               //BUFFER CONVEYOR LEVEL 5 - CONVEYOR 2
               "Control_DB".LCnv_Sys[3].Cnv_Level[5].Cnv2.Inputs.Left := NOT "C3205 - SENSOR CNV LEFT (FWD)";
               "Control_DB".LCnv_Sys[3].Cnv_Level[5].Cnv2.Inputs.Lpd1 := NOT "C3205 - SENSOR CNV LEFT (PALLET DETECT 1)";
               "Control_DB".LCnv_Sys[3].Cnv_Level[5].Cnv2.Inputs.Lpd2 := NOT "C3205 - SENSOR CNV LEFT (PALLET DETECT 2)";
               "Control_DB".LCnv_Sys[3].Cnv_Level[5].Cnv2.Inputs.Right := NOT "C3205 - SENSOR CNV RIGHT (BWD)";
               "Control_DB".LCnv_Sys[3].Cnv_Level[5].Cnv2.Inputs.Rpd1 := NOT "C3205 - SENSOR CNV RIGHT (PALLET DETECT 1)";
               "Control_DB".LCnv_Sys[3].Cnv_Level[5].Cnv2.Inputs.Rpd2 := NOT "C3205 - SENSOR CNV RIGHT (PALLET DETECT 2)";
               "Control_DB".LCnv_Sys[3].Cnv_Level[5].Cnv2.Inputs.Sdetect1 := NOT "C3205 - SHUTTLE IN POSITION 1";
               "Control_DB".LCnv_Sys[3].Cnv_Level[5].Cnv2.Inputs.Sdetect2 := NOT "C3205 - SHUTTLE IN POSITION 2";
               "Control_DB".LCnv_Sys[3].Cnv_Level[5].Cnv2.Safety_Stop_Cnrl.Inputs.DP_Extended := "C3205 - SENSOR SAFETY PIN1 UP";
               "Control_DB".LCnv_Sys[3].Cnv_Level[5].Cnv2.Safety_Stop_Cnrl.Inputs.DP_Retracted := "C3205 - SENSOR SAFETY PIN1 DOWN";

               "Control_DB".LCnv_Sys[3].Cnv_Level[5].Cnv2.Inputs.VFD_Status := "C3205_StatusWord";
               "Control_DB".LCnv_Sys[3].Cnv_Level[5].Cnv2.Inputs.VFD_ActualCurrent := WORD_TO_INT("C3205_ActualCurrent");
               "Control_DB".LCnv_Sys[3].Cnv_Level[5].Cnv2.Inputs.VFD_Speed_Actual := WORD_TO_INT("C3205_ActualSpeed");
               "Control_DB".LCnv_Sys[3].Cnv_Level[5].Cnv2.Inputs.VFD_ActualTorque := WORD_TO_INT("C3205_ActualTorque");
           END_REGION

           REGION LEVEL 6
               //BUFFER CONVEYOR LEVEL 6 - CONVEYOR 1
               "Control_DB".LCnv_Sys[3].Cnv_Level[6].Cnv1.Inputs.Left := NOT "C3106 - SENSOR CNV LEFT (FWD)";
               "Control_DB".LCnv_Sys[3].Cnv_Level[6].Cnv1.Inputs.Lpd1 := NOT "C3106 - SENSOR CNV LEFT (PALLET DETECT 1)";
               "Control_DB".LCnv_Sys[3].Cnv_Level[6].Cnv1.Inputs.Lpd2 := NOT "C3106 - SENSOR CNV LEFT (PALLET DETECT 2)";
               "Control_DB".LCnv_Sys[3].Cnv_Level[6].Cnv1.Inputs.Right := NOT "C3106 - SENSOR CNV RIGHT (BWD)";
               "Control_DB".LCnv_Sys[3].Cnv_Level[6].Cnv1.Inputs.Rpd1 := NOT "C3106 - SENSOR CNV RIGHT (PALLET DETECT 1)";
               "Control_DB".LCnv_Sys[3].Cnv_Level[6].Cnv1.Inputs.Rpd2 := NOT "C3106 - SENSOR CNV RIGHT (PALLET DETECT 2)";
               "Control_DB".LCnv_Sys[3].Cnv_Level[6].Cnv1.Inputs.Sdetect1 := NOT "C3106 - SHUTTLE IN POSITION 1";
               "Control_DB".LCnv_Sys[3].Cnv_Level[6].Cnv1.Inputs.Sdetect2 := NOT "C3106 - SHUTTLE IN POSITION 2";
               "Control_DB".LCnv_Sys[3].Cnv_Level[6].Cnv1.Safety_Stop_Cnrl.Inputs.DP_Extended := "C3106 - SENSOR SAFETY PIN1 UP";
               "Control_DB".LCnv_Sys[3].Cnv_Level[6].Cnv1.Safety_Stop_Cnrl.Inputs.DP_Retracted := "C3106 - SENSOR SAFETY PIN1 DOWN";

               "Control_DB".LCnv_Sys[3].Cnv_Level[6].Cnv1.Inputs.VFD_Status := "C3106_StatusWord";
               "Control_DB".LCnv_Sys[3].Cnv_Level[6].Cnv1.Inputs.VFD_ActualCurrent := WORD_TO_INT("C3106_ActualCurrent");
               "Control_DB".LCnv_Sys[3].Cnv_Level[6].Cnv1.Inputs.VFD_Speed_Actual := WORD_TO_INT("C3106_ActualSpeed");
               "Control_DB".LCnv_Sys[3].Cnv_Level[6].Cnv1.Inputs.VFD_ActualTorque := WORD_TO_INT("C3106_ActualTorque");

               //BUFFER CONVEYOR LEVEL 6 - CONVEYOR 2
               "Control_DB".LCnv_Sys[3].Cnv_Level[6].Cnv2.Inputs.Left := NOT "C3206 - SENSOR CNV LEFT (FWD)";
               "Control_DB".LCnv_Sys[3].Cnv_Level[6].Cnv2.Inputs.Lpd1 := NOT "C3206 - SENSOR CNV LEFT (PALLET DETECT 1)";
               "Control_DB".LCnv_Sys[3].Cnv_Level[6].Cnv2.Inputs.Lpd2 := NOT "C3206 - SENSOR CNV LEFT (PALLET DETECT 2)";
               "Control_DB".LCnv_Sys[3].Cnv_Level[6].Cnv2.Inputs.Right := NOT "C3206 - SENSOR CNV RIGHT (BWD)";
               "Control_DB".LCnv_Sys[3].Cnv_Level[6].Cnv2.Inputs.Rpd1 := NOT "C3206 - SENSOR CNV RIGHT (PALLET DETECT 1)";
               "Control_DB".LCnv_Sys[3].Cnv_Level[6].Cnv2.Inputs.Rpd2 := NOT "C3206 - SENSOR CNV RIGHT (PALLET DETECT 2)";
               "Control_DB".LCnv_Sys[3].Cnv_Level[6].Cnv2.Inputs.Sdetect1 := NOT "C3206 - SHUTTLE IN POSITION 1";
               "Control_DB".LCnv_Sys[3].Cnv_Level[6].Cnv2.Inputs.Sdetect2 := NOT "C3206 - SHUTTLE IN POSITION 2";
               "Control_DB".LCnv_Sys[3].Cnv_Level[6].Cnv2.Safety_Stop_Cnrl.Inputs.DP_Extended := "C3206 - SENSOR SAFETY PIN1 UP";
               "Control_DB".LCnv_Sys[3].Cnv_Level[6].Cnv2.Safety_Stop_Cnrl.Inputs.DP_Retracted := "C3206 - SENSOR SAFETY PIN1 DOWN";

               "Control_DB".LCnv_Sys[3].Cnv_Level[6].Cnv2.Inputs.VFD_Status := "C3206_StatusWord";
               "Control_DB".LCnv_Sys[3].Cnv_Level[6].Cnv2.Inputs.VFD_ActualCurrent := WORD_TO_INT("C3206_ActualCurrent");
               "Control_DB".LCnv_Sys[3].Cnv_Level[6].Cnv2.Inputs.VFD_Speed_Actual := WORD_TO_INT("C3206_ActualSpeed");
               "Control_DB".LCnv_Sys[3].Cnv_Level[6].Cnv2.Inputs.VFD_ActualTorque := WORD_TO_INT("C3206_ActualTorque");
           END_REGION

           REGION LEVEL 7
               //BUFFER CONVEYOR LEVEL 7 - CONVEYOR 1
               "Control_DB".LCnv_Sys[3].Cnv_Level[7].Cnv1.Inputs.Left := NOT "C3107 - SENSOR CNV LEFT (FWD)";
               "Control_DB".LCnv_Sys[3].Cnv_Level[7].Cnv1.Inputs.Lpd1 := NOT "C3107 - SENSOR CNV LEFT (PALLET DETECT 1)";
               "Control_DB".LCnv_Sys[3].Cnv_Level[7].Cnv1.Inputs.Lpd2 := NOT "C3107 - SENSOR CNV LEFT (PALLET DETECT 2)";
               "Control_DB".LCnv_Sys[3].Cnv_Level[7].Cnv1.Inputs.Right := NOT "C3107 - SENSOR CNV RIGHT (BWD)";
               "Control_DB".LCnv_Sys[3].Cnv_Level[7].Cnv1.Inputs.Rpd1 := NOT "C3107 - SENSOR CNV RIGHT (PALLET DETECT 1)";
               "Control_DB".LCnv_Sys[3].Cnv_Level[7].Cnv1.Inputs.Rpd2 := NOT "C3107 - SENSOR CNV RIGHT (PALLET DETECT 2)";
               "Control_DB".LCnv_Sys[3].Cnv_Level[7].Cnv1.Inputs.Sdetect1 := NOT "C3107 - SHUTTLE IN POSITION 1";
               "Control_DB".LCnv_Sys[3].Cnv_Level[7].Cnv1.Inputs.Sdetect2 := NOT "C3107 - SHUTTLE IN POSITION 2";
               "Control_DB".LCnv_Sys[3].Cnv_Level[7].Cnv1.Safety_Stop_Cnrl.Inputs.DP_Extended := "C3107 - SENSOR SAFETY PIN1 UP";
               "Control_DB".LCnv_Sys[3].Cnv_Level[7].Cnv1.Safety_Stop_Cnrl.Inputs.DP_Retracted := "C3107 - SENSOR SAFETY PIN1 DOWN";

               "Control_DB".LCnv_Sys[3].Cnv_Level[7].Cnv1.Inputs.VFD_Status := "C3107_StatusWord";
               "Control_DB".LCnv_Sys[3].Cnv_Level[7].Cnv1.Inputs.VFD_ActualCurrent := WORD_TO_INT("C3107_ActualCurrent");
               "Control_DB".LCnv_Sys[3].Cnv_Level[7].Cnv1.Inputs.VFD_Speed_Actual := WORD_TO_INT("C3107_ActualSpeed");
               "Control_DB".LCnv_Sys[3].Cnv_Level[7].Cnv1.Inputs.VFD_ActualTorque := WORD_TO_INT("C3107_ActualTorque");

               //BUFFER CONVEYOR LEVEL 7 - CONVEYOR 2
               "Control_DB".LCnv_Sys[3].Cnv_Level[7].Cnv2.Inputs.Left := NOT "C3207 - SENSOR CNV LEFT (FWD)";
               "Control_DB".LCnv_Sys[3].Cnv_Level[7].Cnv2.Inputs.Lpd1 := NOT "C3207 - SENSOR CNV LEFT (PALLET DETECT 1)";
               "Control_DB".LCnv_Sys[3].Cnv_Level[7].Cnv2.Inputs.Lpd2 := NOT "C3207 - SENSOR CNV LEFT (PALLET DETECT 2)";
               "Control_DB".LCnv_Sys[3].Cnv_Level[7].Cnv2.Inputs.Right := NOT "C3207 - SENSOR CNV RIGHT (BWD)";
               "Control_DB".LCnv_Sys[3].Cnv_Level[7].Cnv2.Inputs.Rpd1 := NOT "C3207 - SENSOR CNV RIGHT (PALLET DETECT 1)";
               "Control_DB".LCnv_Sys[3].Cnv_Level[7].Cnv2.Inputs.Rpd2 := NOT "C3207 - SENSOR CNV RIGHT (PALLET DETECT 2)";
               "Control_DB".LCnv_Sys[3].Cnv_Level[7].Cnv2.Inputs.Sdetect1 := NOT "C3207 - SHUTTLE IN POSITION 1";
               "Control_DB".LCnv_Sys[3].Cnv_Level[7].Cnv2.Inputs.Sdetect2 := NOT "C3207 - SHUTTLE IN POSITION 2";
               "Control_DB".LCnv_Sys[3].Cnv_Level[7].Cnv2.Safety_Stop_Cnrl.Inputs.DP_Extended := "C3207 - SENSOR SAFETY PIN1 UP";
               "Control_DB".LCnv_Sys[3].Cnv_Level[7].Cnv2.Safety_Stop_Cnrl.Inputs.DP_Retracted := "C3207 - SENSOR SAFETY PIN1 DOWN";

               "Control_DB".LCnv_Sys[3].Cnv_Level[7].Cnv2.Inputs.VFD_Status := "C3207_StatusWord";
               "Control_DB".LCnv_Sys[3].Cnv_Level[7].Cnv2.Inputs.VFD_ActualCurrent := WORD_TO_INT("C3207_ActualCurrent");
               "Control_DB".LCnv_Sys[3].Cnv_Level[7].Cnv2.Inputs.VFD_Speed_Actual := WORD_TO_INT("C3207_ActualSpeed");
               "Control_DB".LCnv_Sys[3].Cnv_Level[7].Cnv2.Inputs.VFD_ActualTorque := WORD_TO_INT("C3207_ActualTorque");
           END_REGION

           REGION LEVEL 8
               //BUFFER CONVEYOR LEVEL 8 - CONVEYOR 1
               "Control_DB".LCnv_Sys[3].Cnv_Level[8].Cnv1.Inputs.Left := NOT "C3108 - SENSOR CNV LEFT (FWD)";
               "Control_DB".LCnv_Sys[3].Cnv_Level[8].Cnv1.Inputs.Lpd1 := NOT "C3108 - SENSOR CNV LEFT (PALLET DETECT 1)";
               "Control_DB".LCnv_Sys[3].Cnv_Level[8].Cnv1.Inputs.Lpd2 := NOT "C3108 - SENSOR CNV LEFT (PALLET DETECT 2)";
               "Control_DB".LCnv_Sys[3].Cnv_Level[8].Cnv1.Inputs.Right := NOT "C3108 - SENSOR CNV RIGHT (BWD)";
               "Control_DB".LCnv_Sys[3].Cnv_Level[8].Cnv1.Inputs.Rpd1 := NOT "C3108 - SENSOR CNV RIGHT (PALLET DETECT 1)";
               "Control_DB".LCnv_Sys[3].Cnv_Level[8].Cnv1.Inputs.Rpd2 := NOT "C3108 - SENSOR CNV RIGHT (PALLET DETECT 2)";
               "Control_DB".LCnv_Sys[3].Cnv_Level[8].Cnv1.Inputs.Sdetect1 := NOT "C3108 - SHUTTLE IN POSITION 1";
               "Control_DB".LCnv_Sys[3].Cnv_Level[8].Cnv1.Inputs.Sdetect2 := NOT "C3108 - SHUTTLE IN POSITION 2";
               "Control_DB".LCnv_Sys[3].Cnv_Level[8].Cnv1.Safety_Stop_Cnrl.Inputs.DP_Extended := "C3108 - SENSOR SAFETY PIN1 UP";
               "Control_DB".LCnv_Sys[3].Cnv_Level[8].Cnv1.Safety_Stop_Cnrl.Inputs.DP_Retracted := "C3108 - SENSOR SAFETY PIN1 DOWN";

               "Control_DB".LCnv_Sys[3].Cnv_Level[8].Cnv1.Inputs.VFD_Status := "C3108_StatusWord";
               "Control_DB".LCnv_Sys[3].Cnv_Level[8].Cnv1.Inputs.VFD_ActualCurrent := WORD_TO_INT("C3108_ActualCurrent");
               "Control_DB".LCnv_Sys[3].Cnv_Level[8].Cnv1.Inputs.VFD_Speed_Actual := WORD_TO_INT("C3108_ActualSpeed");
               "Control_DB".LCnv_Sys[3].Cnv_Level[8].Cnv1.Inputs.VFD_ActualTorque := WORD_TO_INT("C3108_ActualTorque");

               //BUFFER CONVEYOR LEVEL 8 - CONVEYOR 2
               "Control_DB".LCnv_Sys[3].Cnv_Level[8].Cnv2.Inputs.Left := NOT "C3208 - SENSOR CNV LEFT (FWD)";
               "Control_DB".LCnv_Sys[3].Cnv_Level[8].Cnv2.Inputs.Lpd1 := NOT "C3208 - SENSOR CNV LEFT (PALLET DETECT 1)";
               "Control_DB".LCnv_Sys[3].Cnv_Level[8].Cnv2.Inputs.Lpd2 := NOT "C3208 - SENSOR CNV LEFT (PALLET DETECT 2)";
               "Control_DB".LCnv_Sys[3].Cnv_Level[8].Cnv2.Inputs.Right := NOT "C3208 - SENSOR CNV RIGHT (BWD)";
               "Control_DB".LCnv_Sys[3].Cnv_Level[8].Cnv2.Inputs.Rpd1 := NOT "C3208 - SENSOR CNV RIGHT (PALLET DETECT 1)";
               "Control_DB".LCnv_Sys[3].Cnv_Level[8].Cnv2.Inputs.Rpd2 := NOT "C3208 - SENSOR CNV RIGHT (PALLET DETECT 2)";
               "Control_DB".LCnv_Sys[3].Cnv_Level[8].Cnv2.Inputs.Sdetect1 := NOT "C3208 - SHUTTLE IN POSITION 1";
               "Control_DB".LCnv_Sys[3].Cnv_Level[8].Cnv2.Inputs.Sdetect2 := NOT "C3208 - SHUTTLE IN POSITION 2";
               "Control_DB".LCnv_Sys[3].Cnv_Level[8].Cnv2.Safety_Stop_Cnrl.Inputs.DP_Extended := "C3208 - SENSOR SAFETY PIN1 UP";
               "Control_DB".LCnv_Sys[3].Cnv_Level[8].Cnv2.Safety_Stop_Cnrl.Inputs.DP_Retracted := "C3208 - SENSOR SAFETY PIN1 DOWN";

               "Control_DB".LCnv_Sys[3].Cnv_Level[8].Cnv2.Inputs.VFD_Status := "C3208_StatusWord";
               "Control_DB".LCnv_Sys[3].Cnv_Level[8].Cnv2.Inputs.VFD_ActualCurrent := WORD_TO_INT("C3208_ActualCurrent");
               "Control_DB".LCnv_Sys[3].Cnv_Level[8].Cnv2.Inputs.VFD_Speed_Actual := WORD_TO_INT("C3208_ActualSpeed");
               "Control_DB".LCnv_Sys[3].Cnv_Level[8].Cnv2.Inputs.VFD_ActualTorque := WORD_TO_INT("C3208_ActualTorque");
           END_REGION
       END_REGION

       REGION VTD
           "Control_DB".VTD_Sys[3].Inputs.Upper_Overtravel := "OVERTRAVEL UPPER LIMIT - CH1(3)";
           "Control_DB".VTD_Sys[3].Inputs.Upper_limit := "VTD3 UPPER LIMIT";
           "Control_DB".VTD_Sys[3].Inputs.Ultimate_SlowDown := "VTD3 ULTIMATE SLOWDOWN";
           "Control_DB".VTD_Sys[3].Inputs.Ultimate_Creep := "VTD3 ULTIMATE CREEP";
           "Control_DB".VTD_Sys[3].Inputs.Lower_Limit := "VTD3 LOWER LIMIT";
           "Control_DB".VTD_Sys[3].Inputs.Lower_Overtravel := "OVERTRAVEL LOWER LIMIT - CH1(3)";
           "Control_DB".VTD_Sys[3].Inputs.Level_Detect1 := "VTD3 LEVEL DETECT 1";
           "Control_DB".VTD_Sys[3].Inputs.Level_Detect2 := "VTD3 LEVEL DETECT 2";
           "Control_DB".VTD_Sys[3].Inputs.DP1_Extended := "VTD3 DOCKING PINS EXTENDED 1";
           "Control_DB".VTD_Sys[3].Inputs.DP2_Extended := "VTD3 DOCKING PINS EXTENDED 2";
           "Control_DB".VTD_Sys[3].Inputs.DP1_Retracted := "VTD3 DOCKING PINS RETRACTED 1";
           "Control_DB".VTD_Sys[3].Inputs.DP2_Retracted := "VTD3 DOCKING PINS RETRACTED 2";
           "Control_DB".VTD_Sys[3].Inputs.Chain_Slack_1 := NOT "Remote_Panel_DB_3".Chain_Slack_1_Filtered;
           "Control_DB".VTD_Sys[3].Inputs.Chain_Slack_2 := NOT "Remote_Panel_DB_3".Chain_Slack_2_Filtered;
           "Control_DB".VTD_Sys[3].Inputs.Chain_Slack_3 := NOT "Remote_Panel_DB_3".Chain_Slack_3_Filtered;
           "Control_DB".VTD_Sys[3].Inputs.Chain_Slack_4 := NOT "Remote_Panel_DB_3".Chain_Slack_4_Filtered;
           "Control_DB".VTD_Sys[3].Inputs.PushToEnter := "VTD3 PUSH TO ENTER VTD ZONE";
           "Control_DB".VTD_Sys[3].Inputs.PushToExit := "VTD3 PUSH TO EXIT VTD ZONE";

           "Control_DB".VTD_Sys[3].Inputs.VFD_Status := "VTD3_StatusWord";
           "Control_DB".VTD_Sys[3].Inputs.VFD_ActualCurrent := REAL_TO_INT(("VTD3_ActualCurrent" / 10) / 72.5);
           "Control_DB".VTD_Sys[3].Inputs.VFD_Speed_Actual := "VTD3_ActualSpeed";
           "Control_DB".VTD_Sys[3].Inputs.VFD_ActualTorque := WORD_TO_INT("VTD3_ActualTorque");

       END_REGION

       REGION ABSOLUTE ENCODER
           REGION DOCUMENTATION
               //STATUS---------------------------------------------------------------------------------------------------------------------
               //
               //Encoder state word 2 - INPUT WORD 1
               //
               // 15 … 12 Encoder’s Sign-OF-Life (NOT relevant)
               // 11, 10 Reserved
               // 9 Control requested 0 = No control BY the PLC requested 1 = Control BY the PLC requested
               // 8 … 0 Reserved

               //Sensor 1 state word - INPUT WORD 2
               //
               // 15 Encoder error Description 0 = No error 1 = Error The error code is output in G1_XIST2.
               // 14 Park mode activated 0 = Normal operation 1 = Park mode activated Feedback based on G1_STW bit 14: No output OF position data G1_XIST1 AND G1_XIST2
               // 13 Transmission OF absolute position value 0 = No transmission 1 = Position value is output in G1_XIST2
               // 12 Status OF the Preset function (set/shift OF home position executed) 0 = No Preset function active 1 = Preset function is run Feedback based on G1_STW bit 12:  
               // 11 Requirement OF error acknowledgement detected New position value is output in G1_XIST1 AND G1_XIST2. On conclusion OF the Preset function the bit is set TO 0. 0 = No RETURN acknowledgement OF Encoder error 1 = Requirement OF error acknowledgement detected Reaction TO bit 15 in the sensor control word 1 G1_STW is acknowledged (see Table 14)
               // 10 Reserved
               // 9 … 0 NOT supported

               //Position 1 - INPUT WORD 3 AND 4
               // "AE_Position_1_Scaled" := (*SCALE_X(MIN := "Settings_DB".VTD_Settings.VTD_Min_Height,
               //                                   VALUE := *)NORM_X(MIN := 0,
               //                                                   VALUE := (SHL(IN:="AE_Position_1", N:=2) * 0.00228881) (*- "AE_Offset"*),
               //                                                   MAX := 1073741824)(*,
               //                                   MAX := "Settings_DB".VTD_Settings.VTD_Max_Heigh)*);
               // "mm_per_pulse" := 401,5584 / 262144;
               // 
               //CONTROL---------------------------------------------------------------------------------------------------------------------
               //
               //Encoder control word 2 - OUTPUT WORD 1
               //
               // 15 … 12 Master’s Sign-OF-Life (NOT relevant)
               // 10 control BY PLC 0 = No control BY the PLC 1 = Control BY the PLC Enables the PLC BY using control words TO activate / deactivate encoder functions
               // 7 Fault acknowledge Error-buffer handling NOT supported
               // 11, 9, 8, 6 … 0 Reserved
               // "AE_Control_Word_1".%X10 := "AE_PLC_Control";
               // 
               //Sensor 1 control word - OUTPUT WORD 2-------------------------------------------------------------------------------------------
               //
               // 15 Acknowledging a sensor error Description 0 = Encoder error message NOT acknowledged BY PLC 1 = Encoder error message acknowledged BY the PLC
               // 14 Activate park mode 0 = Normal operation 1 = Activate park mode
               // 13 Request FOR the absolute position value 0 = No request 1 = Request BY the master Results in the cyclic output OF the position values in G1_XIST2
               // 12 Activate preset value (see note below) Defines that a configured preset value is used (see section 3.5 on page 24) 0 = Preset value is NOT activated 1 = Preset value is activated
               // 11 Preset mode Defines how a configured preset value is used 0 = Preset value is used as a new absolute value 1 = Preset value is added TO the previous value
               // 10 … 0 Reserved
               // "AE_Control_Word_2".%X15 := "VTD_Reset_HMI_Tags";
               // "AE_Control_Word_2".%X14 := "AE_Activate_ParkMode";
               // "AE_Control_Word_2".%X13 := "AE_Request_ABS_Value";
               // "AE_Control_Word_2".%X12 := "AE_Activate_Preset_Value";
               // "AE_Control_Word_2".%X11 := "AE_Preset_Mode";
           END_REGION

           //STATUS---------------------------------------------------------------------------------------------------------------------
           "Control_DB".VTD_Sys[3].Inputs.AE_Status_2 := "AE_Status_2(3)";
           //Position 1 - INPUT WORD 3 AND 4
           "Control_DB".VTD_Sys[3].Inputs.AE_Position_1 := REAL_TO_DINT(((((*1073741823 - reverse the direction*)
         (SHR(IN := "AE_Position_1(3)", N := 2))) - 31381317) * 0.0015318237304688 (*Mechanical relationship*)- 225511)(*Offset*));

           // Position 2 - INPUT WORD 5 AND 6
           "Control_DB".VTD_Sys[3].Inputs.AE_Position_2 := SHR(IN := "AE_Position_2(3)", N := 2);

           //Speed A - INPUT WORD 7
           "Control_DB".VTD_Sys[3].Inputs.AE_Speed := "AE_Speed(3)";
       END_REGION

       REGION LINEAR ENCODER
           "Control_DB".VTD_Sys[3].Inputs.LE_Position := "LE_X_Unsafe_Position(3)" / 10;
           "Control_DB".VTD_Sys[3].Inputs.LE_Speed := "LE_Speed(3)" * 100;
           "Control_DB".VTD_Sys[3].Inputs.LE_Status := "LE_Status(3)";
           "Control_DB".VTD_Sys[3].Inputs.LE_Warnings := "LE_Warnings(3)";
           REGION DOCUMENTATION
               //STATUS 
               //
               // 0 ERR - Error message (Error code in XP00– XP15); remaining bits = 0, see Error Codes
               // 1 NP - No position information/OUT (XP = 0, YP = 0, SP = 0)
               // 2 WRN - Warnings present, see Warning Module
               // 3 EV - Event present
               // 4 posdetected - Valid position information available

               //WARNINGS
               //
               // 0 WRN01 A code with non-PXV content was found.
               // 1 WRN02 the read head is too close TO the Data Matrix code tape.
               // 2 WRN03 the read head is too far from the Data Matrix code tape.
               // 3 WRN04 Y position too large. The sensor is just before OUT.
               // 4 WRN05 Y position is too small. The sensor is just before OUT.
               // 5 WRN06 the read head is rotated OR tilted in relation TO the Data Matrix code tape.
               // 6 WRN07 Low level OF code contrast.
               // 7 WRN08 Repair tape detected.
               // 8 WRN09 Temperature too high.
               // 9...15 Reserved

               //QUALITY GRADE
               //
               //The quality grades enable constant monitoring of the code tape and the camera along the entire
               //traverse distance. This enables you to detect and act upon potential damage or contamination
               //of the code tape and camera at the earliest stage possible during commissioning and normal
               //operation. As a result, this maximizes the overall functional reliability of your plant, and
               //it means you are able to immediately localize the issue in the case of a fault. Evaluations
               //are made using a scale of 1 to 6. The value 1 is the best possible read quality. A value greater
               //than 3 or worse requires the camera and its path to be inspected. The value 7 signifies "No position"
               //because no code was detected. An evaluation that indicates poor quality as the outcome can be due to
               //a misalignment or incorrect orientation, an incorrect measuring distance, or because the code tape has been affixed incorrectly
           END_REGION
       END_REGION

       REGION SICK BARCODE LECTORS
           IF "Control_DB".VTDBarcode_Station[3].Running AND "SICK_Lector_Control_DB_3".Result <> "Control_DB".VTDBarcode_Station[3].Barcode_Old THEN
               "Control_DB".VTD_Sys[3].Inputs."Barcode 1" := "SICK_Lector_Control_DB_3".Result;
               // "Control_DB".VTD_Control.Inputs."Barcode 2'" := SICK_Barcode_DB".Result;
               // "Control_DB".VTDBarcode_Station[3].Barcode_Old := "SICK_Lector_Control_DB_3".Result;
           ELSE
               "Control_DB".VTD_Sys[3].Inputs."Barcode 1" :=
               "Control_DB".VTD_Sys[3].Inputs."Barcode 2" := '';
           END_IF;

       END_REGION

       REGION VFD HARDWARE ID
           //Buffer conveyors 1
           "Settings_DB".LCnv_Sys[3].Cnv_Level[1].Cnv1.G120_Hardware_ID := "C3101~Drive_1~Standard_telegram_20__PZD-2_6";
           "Settings_DB".LCnv_Sys[3].Cnv_Level[2].Cnv1.G120_Hardware_ID := "C3102~Drive_1~Standard_telegram_20__PZD-2_6";
           "Settings_DB".LCnv_Sys[3].Cnv_Level[3].Cnv1.G120_Hardware_ID := "C3103~Drive_1~Standard_telegram_20__PZD-2_6";
           "Settings_DB".LCnv_Sys[3].Cnv_Level[4].Cnv1.G120_Hardware_ID := "C3104~Drive_1~Standard_telegram_20__PZD-2_6";
           "Settings_DB".LCnv_Sys[3].Cnv_Level[5].Cnv1.G120_Hardware_ID := "C3105~Drive_1~Standard_telegram_20__PZD-2_6";
           "Settings_DB".LCnv_Sys[3].Cnv_Level[6].Cnv1.G120_Hardware_ID := "C3106~Drive_1~Standard_telegram_20__PZD-2_6";
           "Settings_DB".LCnv_Sys[3].Cnv_Level[7].Cnv1.G120_Hardware_ID := "C3107~Drive_1~Standard_telegram_20__PZD-2_6";
           "Settings_DB".LCnv_Sys[3].Cnv_Level[8].Cnv1.G120_Hardware_ID := "C3108~Drive_1~Standard_telegram_20__PZD-2_6";

           //Buffer conveyors 2
           "Settings_DB".LCnv_Sys[3].Cnv_Level[1].Cnv2.G120_Hardware_ID := "C3201~Drive_1~Standard_telegram_20__PZD-2_6";
           "Settings_DB".LCnv_Sys[3].Cnv_Level[2].Cnv2.G120_Hardware_ID := "C3202~Drive_1~Standard_telegram_20__PZD-2_6";
           "Settings_DB".LCnv_Sys[3].Cnv_Level[3].Cnv2.G120_Hardware_ID := "C3203~Drive_1~Standard_telegram_20__PZD-2_6";
           "Settings_DB".LCnv_Sys[3].Cnv_Level[4].Cnv2.G120_Hardware_ID := "C3204~Drive_1~Standard_telegram_20__PZD-2_6";
           "Settings_DB".LCnv_Sys[3].Cnv_Level[5].Cnv2.G120_Hardware_ID := "C3205~Drive_1~Standard_telegram_20__PZD-2_6";
           "Settings_DB".LCnv_Sys[3].Cnv_Level[6].Cnv2.G120_Hardware_ID := "C3206~Drive_1~Standard_telegram_20__PZD-2_6";
           "Settings_DB".LCnv_Sys[3].Cnv_Level[7].Cnv2.G120_Hardware_ID := "C3207~Drive_1~Standard_telegram_20__PZD-2_6";
           "Settings_DB".LCnv_Sys[3].Cnv_Level[8].Cnv2.G120_Hardware_ID := "C3208~Drive_1~Standard_telegram_20__PZD-2_6";

           //Extractor conveyor
           "Settings_DB".ECnv_Sys[3].G120_Hardware_ID := "CVTD_3~Drive_1~Standard_telegram_20__PZD-2_6";

           //VTD
           "Settings_DB".VTD_Sys[3].G120_Hardware_ID := "VTD_3~DO_VECTOR_1~Standard_telegram_20__PZD-2_6";
       END_REGION
   END_REGION

   REGION SYSTEM 4
       REGION EXTRACTOR CONVEYOR
           "Control_DB".ECnv_Sys[4].Inputs.Left := "CVTD4 SENSOR CONVEYOR LEFT (FWD)";
           "Control_DB".ECnv_Sys[4].Inputs.Lpd1 := "CVTD4 SENSOR CONVEYOR LEFT (PALLET DETECT 1)";
           "Control_DB".ECnv_Sys[4].Inputs.Center := "CVTD4 SENSOR CONVEYOR CENTER";
           "Control_DB".ECnv_Sys[4].Inputs.Right := "CVTD4 SENSOR CONVEYOR RIGHT (BWD)";
           "Control_DB".ECnv_Sys[4].Inputs.Rpd1 := "CVTD4 SENSOR CONVEYOR RIGHT (PALLET DETECT 1)";

           "T_OH_Left_4".TOF(IN := "CVTD4 OVERHANG LEFT" OR NOT "Control_DB".VTD_Sys[4].Running,
                             PT := T#200ms);
           "Control_DB".ECnv_Sys[4].Inputs.Overhang_Left := "T_OH_Left_4".Q;

           "I_OH_Right_4".TOF(IN := "CVTD4 OVERHANG RIGHT" OR NOT "Control_DB".VTD_Sys[4].Running,
                              PT := T#200ms);
           "Control_DB".ECnv_Sys[4].Inputs.Overhang_Right := "I_OH_Right_4".Q;

           "Control_DB".ECnv_Sys[4].Inputs.VFD_Status := "CVTD4_StatusWord";
           "Control_DB".ECnv_Sys[4].Inputs.VFD_ActualCurrent := WORD_TO_INT("CVTD4_ActualCurrent");
           "Control_DB".ECnv_Sys[4].Inputs.VFD_Speed_Actual := WORD_TO_INT("CVTD4_ActualSpeed");
           "Control_DB".ECnv_Sys[4].Inputs.VFD_ActualTorque := WORD_TO_INT("CVTD4_ActualTorque");
       END_REGION

       REGION BUFFER CONVEYORS
           REGION LEVEL 1
               //BUFFER CONVEYOR LEVEL 1 - CONVEYOR 1
               "Control_DB".LCnv_Sys[4].Cnv_Level[1].Cnv1.Inputs.Left := NOT "C4101 - SENSOR CNV LEFT (FWD)";
               "Control_DB".LCnv_Sys[4].Cnv_Level[1].Cnv1.Inputs.Lpd1 := NOT "C4101 - SENSOR CNV LEFT (PALLET DETECT 1)";
               "Control_DB".LCnv_Sys[4].Cnv_Level[1].Cnv1.Inputs.Lpd2 := NOT "C4101 - SENSOR CNV LEFT (PALLET DETECT 2)";
               "Control_DB".LCnv_Sys[4].Cnv_Level[1].Cnv1.Inputs.Right := NOT "C4101 - SENSOR CNV RIGHT (BWD)";
               "Control_DB".LCnv_Sys[4].Cnv_Level[1].Cnv1.Inputs.Rpd1 := NOT "C4101 - SENSOR CNV RIGHT (PALLET DETECT 1)";
               "Control_DB".LCnv_Sys[4].Cnv_Level[1].Cnv1.Inputs.Rpd2 := NOT "C4101 - SENSOR CNV RIGHT (PALLET DETECT 2)";
               "Control_DB".LCnv_Sys[4].Cnv_Level[1].Cnv1.Inputs.Sdetect1 := NOT "C4101 - SHUTTLE IN POSITION 1";
               "Control_DB".LCnv_Sys[4].Cnv_Level[1].Cnv1.Inputs.Sdetect2 := NOT "C4101 - SHUTTLE IN POSITION 2";
               "Control_DB".LCnv_Sys[4].Cnv_Level[1].Cnv1.Safety_Stop_Cnrl.Inputs.DP_Extended := "C4101 - SENSOR SAFETY PIN1 UP";
               "Control_DB".LCnv_Sys[4].Cnv_Level[1].Cnv1.Safety_Stop_Cnrl.Inputs.DP_Retracted := "C4101 - SENSOR SAFETY PIN1 DOWN";

               "Control_DB".LCnv_Sys[4].Cnv_Level[1].Cnv1.Inputs.VFD_Status := "C4101_StatusWord";
               "Control_DB".LCnv_Sys[4].Cnv_Level[1].Cnv1.Inputs.VFD_ActualCurrent := WORD_TO_INT("C4101_ActualCurrent");
               "Control_DB".LCnv_Sys[4].Cnv_Level[1].Cnv1.Inputs.VFD_Speed_Actual := WORD_TO_INT("C4101_ActualSpeed");
               "Control_DB".LCnv_Sys[4].Cnv_Level[1].Cnv1.Inputs.VFD_ActualTorque := WORD_TO_INT("C4101_ActualTorque");
           END_REGION

           REGION LEVEL 2
               //BUFFER CONVEYOR LEVEL 2 - CONVEYOR 1
               "Control_DB".LCnv_Sys[4].Cnv_Level[2].Cnv1.Inputs.Left := NOT "C4102 - SENSOR CNV LEFT (FWD)";
               "Control_DB".LCnv_Sys[4].Cnv_Level[2].Cnv1.Inputs.Lpd1 := NOT "C4102 - SENSOR CNV LEFT (PALLET DETECT 1)";
               "Control_DB".LCnv_Sys[4].Cnv_Level[2].Cnv1.Inputs.Lpd2 := NOT "C4102 - SENSOR CNV LEFT (PALLET DETECT 2)";
               "Control_DB".LCnv_Sys[4].Cnv_Level[2].Cnv1.Inputs.Right := NOT "C4102 - SENSOR CNV RIGHT (BWD)";
               "Control_DB".LCnv_Sys[4].Cnv_Level[2].Cnv1.Inputs.Rpd1 := NOT "C4102 - SENSOR CNV RIGHT (PALLET DETECT 1)";
               "Control_DB".LCnv_Sys[4].Cnv_Level[2].Cnv1.Inputs.Rpd2 := NOT "C4102 - SENSOR CNV RIGHT (PALLET DETECT 2)";
               "Control_DB".LCnv_Sys[4].Cnv_Level[2].Cnv1.Inputs.Sdetect1 := NOT "C4102 - SHUTTLE IN POSITION 1";
               "Control_DB".LCnv_Sys[4].Cnv_Level[2].Cnv1.Inputs.Sdetect2 := NOT "C4102 - SHUTTLE IN POSITION 2";
               "Control_DB".LCnv_Sys[4].Cnv_Level[2].Cnv1.Safety_Stop_Cnrl.Inputs.DP_Extended := "C4102 - SENSOR SAFETY PIN1 UP";
               "Control_DB".LCnv_Sys[4].Cnv_Level[2].Cnv1.Safety_Stop_Cnrl.Inputs.DP_Retracted := "C4102 - SENSOR SAFETY PIN1 DOWN";

               "Control_DB".LCnv_Sys[4].Cnv_Level[2].Cnv1.Inputs.VFD_Status := "C4102_StatusWord";
               "Control_DB".LCnv_Sys[4].Cnv_Level[2].Cnv1.Inputs.VFD_ActualCurrent := WORD_TO_INT("C4102_ActualCurrent");
               "Control_DB".LCnv_Sys[4].Cnv_Level[2].Cnv1.Inputs.VFD_Speed_Actual := WORD_TO_INT("C4102_ActualSpeed");
               "Control_DB".LCnv_Sys[4].Cnv_Level[2].Cnv1.Inputs.VFD_ActualTorque := WORD_TO_INT("C4102_ActualTorque");
           END_REGION

           REGION LEVEL 3
               //BUFFER CONVEYOR LEVEL 3 - CONVEYOR 1
               "Control_DB".LCnv_Sys[4].Cnv_Level[3].Cnv1.Inputs.Left := NOT "C4103 - SENSOR CNV LEFT (FWD)";
               "Control_DB".LCnv_Sys[4].Cnv_Level[3].Cnv1.Inputs.Lpd1 := NOT "C4103 - SENSOR CNV LEFT (PALLET DETECT 1)";
               "Control_DB".LCnv_Sys[4].Cnv_Level[3].Cnv1.Inputs.Lpd2 := NOT "C4103 - SENSOR CNV LEFT (PALLET DETECT 2)";
               "Control_DB".LCnv_Sys[4].Cnv_Level[3].Cnv1.Inputs.Right := NOT "C4103 - SENSOR CNV RIGHT (BWD)";
               "Control_DB".LCnv_Sys[4].Cnv_Level[3].Cnv1.Inputs.Rpd1 := NOT "C4103 - SENSOR CNV RIGHT (PALLET DETECT 1)";
               "Control_DB".LCnv_Sys[4].Cnv_Level[3].Cnv1.Inputs.Rpd2 := NOT "C4103 - SENSOR CNV RIGHT (PALLET DETECT 2)";
               "Control_DB".LCnv_Sys[4].Cnv_Level[3].Cnv1.Inputs.Sdetect1 := NOT "C4103 - SHUTTLE IN POSITION 1";
               "Control_DB".LCnv_Sys[4].Cnv_Level[3].Cnv1.Inputs.Sdetect2 := NOT "C4103 - SHUTTLE IN POSITION 2";
               "Control_DB".LCnv_Sys[4].Cnv_Level[3].Cnv1.Safety_Stop_Cnrl.Inputs.DP_Extended := "C4103 - SENSOR SAFETY PIN1 UP";
               "Control_DB".LCnv_Sys[4].Cnv_Level[3].Cnv1.Safety_Stop_Cnrl.Inputs.DP_Retracted := "C4103 - SENSOR SAFETY PIN1 DOWN";

               "Control_DB".LCnv_Sys[4].Cnv_Level[3].Cnv1.Inputs.VFD_Status := "C4103_StatusWord";
               "Control_DB".LCnv_Sys[4].Cnv_Level[3].Cnv1.Inputs.VFD_ActualCurrent := WORD_TO_INT("C4103_ActualCurrent");
               "Control_DB".LCnv_Sys[4].Cnv_Level[3].Cnv1.Inputs.VFD_Speed_Actual := WORD_TO_INT("C4103_ActualSpeed");
               "Control_DB".LCnv_Sys[4].Cnv_Level[3].Cnv1.Inputs.VFD_ActualTorque := WORD_TO_INT("C4103_ActualTorque");
           END_REGION

           REGION LEVEL 4
               //BUFFER CONVEYOR LEVEL 4 - CONVEYOR 1
               "Control_DB".LCnv_Sys[4].Cnv_Level[4].Cnv1.Inputs.Left := NOT "C4104 - SENSOR CNV LEFT (FWD)";
               "Control_DB".LCnv_Sys[4].Cnv_Level[4].Cnv1.Inputs.Lpd1 := NOT "C4104 - SENSOR CNV LEFT (PALLET DETECT 1)";
               "Control_DB".LCnv_Sys[4].Cnv_Level[4].Cnv1.Inputs.Lpd2 := NOT "C4104 - SENSOR CNV LEFT (PALLET DETECT 2)";
               "Control_DB".LCnv_Sys[4].Cnv_Level[4].Cnv1.Inputs.Right := NOT "C4104 - SENSOR CNV RIGHT (BWD)";
               "Control_DB".LCnv_Sys[4].Cnv_Level[4].Cnv1.Inputs.Rpd1 := NOT "C4104 - SENSOR CNV RIGHT (PALLET DETECT 1)";
               "Control_DB".LCnv_Sys[4].Cnv_Level[4].Cnv1.Inputs.Rpd2 := NOT "C4104 - SENSOR CNV RIGHT (PALLET DETECT 2)";
               "Control_DB".LCnv_Sys[4].Cnv_Level[4].Cnv1.Inputs.Sdetect1 := NOT "C4104 - SHUTTLE IN POSITION 1";
               "Control_DB".LCnv_Sys[4].Cnv_Level[4].Cnv1.Inputs.Sdetect2 := NOT "C4104 - SHUTTLE IN POSITION 2";
               "Control_DB".LCnv_Sys[4].Cnv_Level[4].Cnv1.Safety_Stop_Cnrl.Inputs.DP_Extended := "C4104 - SENSOR SAFETY PIN1 UP";
               "Control_DB".LCnv_Sys[4].Cnv_Level[4].Cnv1.Safety_Stop_Cnrl.Inputs.DP_Retracted := "C4104 - SENSOR SAFETY PIN1 DOWN";

               "Control_DB".LCnv_Sys[4].Cnv_Level[4].Cnv1.Inputs.VFD_Status := "C4104_StatusWord";
               "Control_DB".LCnv_Sys[4].Cnv_Level[4].Cnv1.Inputs.VFD_ActualCurrent := WORD_TO_INT("C4104_ActualCurrent");
               "Control_DB".LCnv_Sys[4].Cnv_Level[4].Cnv1.Inputs.VFD_Speed_Actual := WORD_TO_INT("C4104_ActualSpeed");
               "Control_DB".LCnv_Sys[4].Cnv_Level[4].Cnv1.Inputs.VFD_ActualTorque := WORD_TO_INT("C4104_ActualTorque");

           END_REGION

           REGION LEVEL 5
               //BUFFER CONVEYOR LEVEL 5 - CONVEYOR 1
               "Control_DB".LCnv_Sys[4].Cnv_Level[5].Cnv1.Inputs.Left := NOT "C4105 - SENSOR CNV LEFT (FWD)";
               "Control_DB".LCnv_Sys[4].Cnv_Level[5].Cnv1.Inputs.Lpd1 := NOT "C4105 - SENSOR CNV LEFT (PALLET DETECT 1)";
               "Control_DB".LCnv_Sys[4].Cnv_Level[5].Cnv1.Inputs.Lpd2 := NOT "C4105 - SENSOR CNV LEFT (PALLET DETECT 2)";
               "Control_DB".LCnv_Sys[4].Cnv_Level[5].Cnv1.Inputs.Right := NOT "C4105 - SENSOR CNV RIGHT (BWD)";
               "Control_DB".LCnv_Sys[4].Cnv_Level[5].Cnv1.Inputs.Rpd1 := NOT "C4105 - SENSOR CNV RIGHT (PALLET DETECT 1)";
               "Control_DB".LCnv_Sys[4].Cnv_Level[5].Cnv1.Inputs.Rpd2 := NOT "C4105 - SENSOR CNV RIGHT (PALLET DETECT 2)";
               "Control_DB".LCnv_Sys[4].Cnv_Level[5].Cnv1.Inputs.Sdetect1 := NOT "C4105 - SHUTTLE IN POSITION 1";
               "Control_DB".LCnv_Sys[4].Cnv_Level[5].Cnv1.Inputs.Sdetect2 := NOT "C4105 - SHUTTLE IN POSITION 2";
               "Control_DB".LCnv_Sys[4].Cnv_Level[5].Cnv1.Safety_Stop_Cnrl.Inputs.DP_Extended := "C4105 - SENSOR SAFETY PIN1 UP";
               "Control_DB".LCnv_Sys[4].Cnv_Level[5].Cnv1.Safety_Stop_Cnrl.Inputs.DP_Retracted := "C4105 - SENSOR SAFETY PIN1 DOWN";

               "Control_DB".LCnv_Sys[4].Cnv_Level[5].Cnv1.Inputs.VFD_Status := "C4105_StatusWord";
               "Control_DB".LCnv_Sys[4].Cnv_Level[5].Cnv1.Inputs.VFD_ActualCurrent := WORD_TO_INT("C4105_ActualCurrent");
               "Control_DB".LCnv_Sys[4].Cnv_Level[5].Cnv1.Inputs.VFD_Speed_Actual := WORD_TO_INT("C4105_ActualSpeed");
               "Control_DB".LCnv_Sys[4].Cnv_Level[5].Cnv1.Inputs.VFD_ActualTorque := WORD_TO_INT("C4105_ActualTorque");
           END_REGION

           REGION LEVEL 6
               //BUFFER CONVEYOR LEVEL 6 - CONVEYOR 1
               "Control_DB".LCnv_Sys[4].Cnv_Level[6].Cnv1.Inputs.Left := NOT "C4106 - SENSOR CNV LEFT (FWD)";
               "Control_DB".LCnv_Sys[4].Cnv_Level[6].Cnv1.Inputs.Lpd1 := NOT "C4106 - SENSOR CNV LEFT (PALLET DETECT 1)";
               "Control_DB".LCnv_Sys[4].Cnv_Level[6].Cnv1.Inputs.Lpd2 := NOT "C4106 - SENSOR CNV LEFT (PALLET DETECT 2)";
               "Control_DB".LCnv_Sys[4].Cnv_Level[6].Cnv1.Inputs.Right := NOT "C4106 - SENSOR CNV RIGHT (BWD)";
               "Control_DB".LCnv_Sys[4].Cnv_Level[6].Cnv1.Inputs.Rpd1 := NOT "C4106 - SENSOR CNV RIGHT (PALLET DETECT 1)";
               "Control_DB".LCnv_Sys[4].Cnv_Level[6].Cnv1.Inputs.Rpd2 := NOT "C4106 - SENSOR CNV RIGHT (PALLET DETECT 2)";
               "Control_DB".LCnv_Sys[4].Cnv_Level[6].Cnv1.Inputs.Sdetect1 := NOT "C4106 - SHUTTLE IN POSITION 1";
               "Control_DB".LCnv_Sys[4].Cnv_Level[6].Cnv1.Inputs.Sdetect2 := NOT "C4106 - SHUTTLE IN POSITION 2";
               "Control_DB".LCnv_Sys[4].Cnv_Level[6].Cnv1.Safety_Stop_Cnrl.Inputs.DP_Extended := "C4106 - SENSOR SAFETY PIN1 UP";
               "Control_DB".LCnv_Sys[4].Cnv_Level[6].Cnv1.Safety_Stop_Cnrl.Inputs.DP_Retracted := "C4106 - SENSOR SAFETY PIN1 DOWN";

               "Control_DB".LCnv_Sys[4].Cnv_Level[6].Cnv1.Inputs.VFD_Status := "C4106_StatusWord";
               "Control_DB".LCnv_Sys[4].Cnv_Level[6].Cnv1.Inputs.VFD_ActualCurrent := WORD_TO_INT("C4106_ActualCurrent");
               "Control_DB".LCnv_Sys[4].Cnv_Level[6].Cnv1.Inputs.VFD_Speed_Actual := WORD_TO_INT("C4106_ActualSpeed");
               "Control_DB".LCnv_Sys[4].Cnv_Level[6].Cnv1.Inputs.VFD_ActualTorque := WORD_TO_INT("C4106_ActualTorque");
           END_REGION

           REGION LEVEL 7
               //BUFFER CONVEYOR LEVEL 7 - CONVEYOR 1
               "Control_DB".LCnv_Sys[4].Cnv_Level[7].Cnv1.Inputs.Left := NOT "C4107 - SENSOR CNV LEFT (FWD)";
               "Control_DB".LCnv_Sys[4].Cnv_Level[7].Cnv1.Inputs.Lpd1 := NOT "C4107 - SENSOR CNV LEFT (PALLET DETECT 1)";
               "Control_DB".LCnv_Sys[4].Cnv_Level[7].Cnv1.Inputs.Lpd2 := NOT "C4107 - SENSOR CNV LEFT (PALLET DETECT 2)";
               "Control_DB".LCnv_Sys[4].Cnv_Level[7].Cnv1.Inputs.Right := NOT "C4107 - SENSOR CNV RIGHT (BWD)";
               "Control_DB".LCnv_Sys[4].Cnv_Level[7].Cnv1.Inputs.Rpd1 := NOT "C4107 - SENSOR CNV RIGHT (PALLET DETECT 1)";
               "Control_DB".LCnv_Sys[4].Cnv_Level[7].Cnv1.Inputs.Rpd2 := NOT "C4107 - SENSOR CNV RIGHT (PALLET DETECT 2)";
               "Control_DB".LCnv_Sys[4].Cnv_Level[7].Cnv1.Inputs.Sdetect1 := NOT "C4107 - SHUTTLE IN POSITION 1";
               "Control_DB".LCnv_Sys[4].Cnv_Level[7].Cnv1.Inputs.Sdetect2 := NOT "C4107 - SHUTTLE IN POSITION 2";
               "Control_DB".LCnv_Sys[4].Cnv_Level[7].Cnv1.Safety_Stop_Cnrl.Inputs.DP_Extended := "C4107 - SENSOR SAFETY PIN1 UP";
               "Control_DB".LCnv_Sys[4].Cnv_Level[7].Cnv1.Safety_Stop_Cnrl.Inputs.DP_Retracted := "C4107 - SENSOR SAFETY PIN1 DOWN";

               "Control_DB".LCnv_Sys[4].Cnv_Level[7].Cnv1.Inputs.VFD_Status := "C4107_StatusWord";
               "Control_DB".LCnv_Sys[4].Cnv_Level[7].Cnv1.Inputs.VFD_ActualCurrent := WORD_TO_INT("C4107_ActualCurrent");
               "Control_DB".LCnv_Sys[4].Cnv_Level[7].Cnv1.Inputs.VFD_Speed_Actual := WORD_TO_INT("C4107_ActualSpeed");
               "Control_DB".LCnv_Sys[4].Cnv_Level[7].Cnv1.Inputs.VFD_ActualTorque := WORD_TO_INT("C4107_ActualTorque");
           END_REGION

           REGION LEVEL 8
               //BUFFER CONVEYOR LEVEL 8 - CONVEYOR 1
               "Control_DB".LCnv_Sys[4].Cnv_Level[8].Cnv1.Inputs.Left := NOT "C4108 - SENSOR CNV LEFT (FWD)";
               "Control_DB".LCnv_Sys[4].Cnv_Level[8].Cnv1.Inputs.Lpd1 := NOT "C4108 - SENSOR CNV LEFT (PALLET DETECT 1)";
               "Control_DB".LCnv_Sys[4].Cnv_Level[8].Cnv1.Inputs.Lpd2 := NOT "C4108 - SENSOR CNV LEFT (PALLET DETECT 2)";
               "Control_DB".LCnv_Sys[4].Cnv_Level[8].Cnv1.Inputs.Right := NOT "C4108 - SENSOR CNV RIGHT (BWD)";
               "Control_DB".LCnv_Sys[4].Cnv_Level[8].Cnv1.Inputs.Rpd1 := NOT "C4108 - SENSOR CNV RIGHT (PALLET DETECT 1)";
               "Control_DB".LCnv_Sys[4].Cnv_Level[8].Cnv1.Inputs.Rpd2 := NOT "C4108 - SENSOR CNV RIGHT (PALLET DETECT 2)";
               "Control_DB".LCnv_Sys[4].Cnv_Level[8].Cnv1.Inputs.Sdetect1 := NOT "C4108 - SHUTTLE IN POSITION 1";
               "Control_DB".LCnv_Sys[4].Cnv_Level[8].Cnv1.Inputs.Sdetect2 := NOT "C4108 - SHUTTLE IN POSITION 2";
               "Control_DB".LCnv_Sys[4].Cnv_Level[8].Cnv1.Safety_Stop_Cnrl.Inputs.DP_Extended := "C4108 - SENSOR SAFETY PIN1 UP";
               "Control_DB".LCnv_Sys[4].Cnv_Level[8].Cnv1.Safety_Stop_Cnrl.Inputs.DP_Retracted := "C4108 - SENSOR SAFETY PIN1 DOWN";

               "Control_DB".LCnv_Sys[4].Cnv_Level[8].Cnv1.Inputs.VFD_Status := "C4108_StatusWord";
               "Control_DB".LCnv_Sys[4].Cnv_Level[8].Cnv1.Inputs.VFD_ActualCurrent := WORD_TO_INT("C4108_ActualCurrent");
               "Control_DB".LCnv_Sys[4].Cnv_Level[8].Cnv1.Inputs.VFD_Speed_Actual := WORD_TO_INT("C4108_ActualSpeed");
               "Control_DB".LCnv_Sys[4].Cnv_Level[8].Cnv1.Inputs.VFD_ActualTorque := WORD_TO_INT("C4108_ActualTorque");
           END_REGION
       END_REGION

       REGION VTD
           "Control_DB".VTD_Sys[4].Inputs.Upper_Overtravel := "OVERTRAVEL UPPER LIMIT - CH1(4)";
           "Control_DB".VTD_Sys[4].Inputs.Upper_limit := "VTD4 UPPER LIMIT";
           "Control_DB".VTD_Sys[4].Inputs.Ultimate_SlowDown := "VTD4 ULTIMATE SLOWDOWN";
           "Control_DB".VTD_Sys[4].Inputs.Ultimate_Creep := "VTD4 ULTIMATE CREEP";
           "Control_DB".VTD_Sys[4].Inputs.Lower_Limit := "VTD4 LOWER LIMIT";
           "Control_DB".VTD_Sys[4].Inputs.Lower_Overtravel := "OVERTRAVEL LOWER LIMIT - CH1(4)";
           "Control_DB".VTD_Sys[4].Inputs.Level_Detect1 := "VTD4 LEVEL DETECT 1";
           "Control_DB".VTD_Sys[4].Inputs.Level_Detect2 := "VTD4 LEVEL DETECT 2";
           "Control_DB".VTD_Sys[4].Inputs.DP1_Extended := "VTD4 DOCKING PINS 1 EXTENDED";
           "Control_DB".VTD_Sys[4].Inputs.DP2_Extended := "VTD4 DOCKING PINS 2 EXTENDED";
           "Control_DB".VTD_Sys[4].Inputs.DP1_Retracted := "VTD4 DOCKING PINS 1 RETRACTED";
           "Control_DB".VTD_Sys[4].Inputs.DP2_Retracted := "VTD4 DOCKING PINS 2 RETRACTED";
           "Control_DB".VTD_Sys[4].Inputs.Chain_Slack_1 := NOT "Remote_Panel_DB_4".Chain_Slack_1_Filtered;
           "Control_DB".VTD_Sys[4].Inputs.Chain_Slack_2 := NOT "Remote_Panel_DB_4".Chain_Slack_2_Filtered;
           "Control_DB".VTD_Sys[4].Inputs.Chain_Slack_3 := NOT "Remote_Panel_DB_4".Chain_Slack_3_Filtered;
           "Control_DB".VTD_Sys[4].Inputs.Chain_Slack_4 := NOT "Remote_Panel_DB_4".Chain_Slack_4_Filtered;
           "Control_DB".VTD_Sys[4].Inputs.PushToEnter := "VTD4 PUSH TO ENTER VTD ZONE";
           "Control_DB".VTD_Sys[4].Inputs.PushToExit := "VTD4 PUSH TO EXIT VTD ZONE";
           "Control_DB".VTD_Sys[4].Inputs.VFD_Status := "VTD4_StatusWord";
           "Control_DB".VTD_Sys[4].Inputs.VFD_ActualCurrent := REAL_TO_INT(("VTD4_ActualCurrent" / 10) / 72.5);
           "Control_DB".VTD_Sys[4].Inputs.VFD_Speed_Actual := "VTD4_ActualSpeed";
           "Control_DB".VTD_Sys[4].Inputs.VFD_ActualTorque := WORD_TO_INT("VTD4_ActualTorque");

       END_REGION

       REGION ABSOLUTE ENCODER
           REGION DOCUMENTATION
               //STATUS---------------------------------------------------------------------------------------------------------------------
               //
               //Encoder state word 2 - INPUT WORD 1
               //
               // 15 … 12 Encoder’s Sign-OF-Life (NOT relevant)
               // 11, 10 Reserved
               // 9 Control requested 0 = No control BY the PLC requested 1 = Control BY the PLC requested
               // 8 … 0 Reserved

               //Sensor 1 state word - INPUT WORD 2
               //
               // 15 Encoder error Description 0 = No error 1 = Error The error code is output in G1_XIST2.
               // 14 Park mode activated 0 = Normal operation 1 = Park mode activated Feedback based on G1_STW bit 14: No output OF position data G1_XIST1 AND G1_XIST2
               // 13 Transmission OF absolute position value 0 = No transmission 1 = Position value is output in G1_XIST2
               // 12 Status OF the Preset function (set/shift OF home position executed) 0 = No Preset function active 1 = Preset function is run Feedback based on G1_STW bit 12:  
               // 11 Requirement OF error acknowledgement detected New position value is output in G1_XIST1 AND G1_XIST2. On conclusion OF the Preset function the bit is set TO 0. 0 = No RETURN acknowledgement OF Encoder error 1 = Requirement OF error acknowledgement detected Reaction TO bit 15 in the sensor control word 1 G1_STW is acknowledged (see Table 14)
               // 10 Reserved
               // 9 … 0 NOT supported

               //Position 1 - INPUT WORD 3 AND 4
               // "AE_Position_1_Scaled" := (*SCALE_X(MIN := "Settings_DB".VTD_Settings.VTD_Min_Height,
               //                                   VALUE := *)NORM_X(MIN := 0,
               //                                                   VALUE := (SHL(IN:="AE_Position_1", N:=2) * 0.00228881) (*- "AE_Offset"*),
               //                                                   MAX := 1073741824)(*,
               //                                   MAX := "Settings_DB".VTD_Settings.VTD_Max_Heigh)*);
               // "mm_per_pulse" := 401,5584 / 262144;
               // 
               //CONTROL---------------------------------------------------------------------------------------------------------------------
               //
               //Encoder control word 2 - OUTPUT WORD 1
               //
               // 15 … 12 Master’s Sign-OF-Life (NOT relevant)
               // 10 control BY PLC 0 = No control BY the PLC 1 = Control BY the PLC Enables the PLC BY using control words TO activate / deactivate encoder functions
               // 7 Fault acknowledge Error-buffer handling NOT supported
               // 11, 9, 8, 6 … 0 Reserved
               // "AE_Control_Word_1".%X10 := "AE_PLC_Control";
               // 
               //Sensor 1 control word - OUTPUT WORD 2-------------------------------------------------------------------------------------------
               //
               // 15 Acknowledging a sensor error Description 0 = Encoder error message NOT acknowledged BY PLC 1 = Encoder error message acknowledged BY the PLC
               // 14 Activate park mode 0 = Normal operation 1 = Activate park mode
               // 13 Request FOR the absolute position value 0 = No request 1 = Request BY the master Results in the cyclic output OF the position values in G1_XIST2
               // 12 Activate preset value (see note below) Defines that a configured preset value is used (see section 3.5 on page 24) 0 = Preset value is NOT activated 1 = Preset value is activated
               // 11 Preset mode Defines how a configured preset value is used 0 = Preset value is used as a new absolute value 1 = Preset value is added TO the previous value
               // 10 … 0 Reserved
               // "AE_Control_Word_2".%X15 := "VTD_Reset_HMI_Tags";
               // "AE_Control_Word_2".%X14 := "AE_Activate_ParkMode";
               // "AE_Control_Word_2".%X13 := "AE_Request_ABS_Value";
               // "AE_Control_Word_2".%X12 := "AE_Activate_Preset_Value";
               // "AE_Control_Word_2".%X11 := "AE_Preset_Mode";
           END_REGION

           //STATUS---------------------------------------------------------------------------------------------------------------------
           "Control_DB".VTD_Sys[4].Inputs.AE_Status_2 := "AE_Status_2(4)";
           //Position 1 - INPUT WORD 3 AND 4
           "Control_DB".VTD_Sys[4].Inputs.AE_Position_1 := REAL_TO_DINT((((1073741823 - (*reverse the direction*)
    (SHR(IN := "AE_Position_1(4)", N := 2))) - 31381317) * 0.0015318237304688 (*Mechanical relationship*)- 935884) (*Offset*));

           // Position 2 - INPUT WORD 5 AND 6
           "Control_DB".VTD_Sys[4].Inputs.AE_Position_2 := SHR(IN := "AE_Position_2(4)", N := 2);

           //Speed A - INPUT WORD 7
           "Control_DB".VTD_Sys[4].Inputs.AE_Speed := "AE_Speed(4)";
       END_REGION

       REGION LINEAR ENCODER
           "Control_DB".VTD_Sys[4].Inputs.LE_Position := "LE_X_Unsafe_Position(4)" / 10;
           "Control_DB".VTD_Sys[4].Inputs.LE_Speed := "LE_Speed(4)" * 100;
           "Control_DB".VTD_Sys[4].Inputs.LE_Status := "LE_Status(4)";
           "Control_DB".VTD_Sys[4].Inputs.LE_Warnings := "LE_Warnings(4)";
           REGION DOCUMENTATION
               //STATUS 
               //
               // 0 ERR - Error message (Error code in XP00– XP15); remaining bits = 0, see Error Codes
               // 1 NP - No position information/OUT (XP = 0, YP = 0, SP = 0)
               // 2 WRN - Warnings present, see Warning Module
               // 3 EV - Event present
               // 4 posdetected - Valid position information available

               //WARNINGS
               //
               // 0 WRN01 A code with non-PXV content was found.
               // 1 WRN02 the read head is too close TO the Data Matrix code tape.
               // 2 WRN03 the read head is too far from the Data Matrix code tape.
               // 3 WRN04 Y position too large. The sensor is just before OUT.
               // 4 WRN05 Y position is too small. The sensor is just before OUT.
               // 5 WRN06 the read head is rotated OR tilted in relation TO the Data Matrix code tape.
               // 6 WRN07 Low level OF code contrast.
               // 7 WRN08 Repair tape detected.
               // 8 WRN09 Temperature too high.
               // 9...15 Reserved

               //QUALITY GRADE
               //
               //The quality grades enable constant monitoring of the code tape and the camera along the entire
               //traverse distance. This enables you to detect and act upon potential damage or contamination
               //of the code tape and camera at the earliest stage possible during commissioning and normal
               //operation. As a result, this maximizes the overall functional reliability of your plant, and
               //it means you are able to immediately localize the issue in the case of a fault. Evaluations
               //are made using a scale of 1 to 6. The value 1 is the best possible read quality. A value greater
               //than 3 or worse requires the camera and its path to be inspected. The value 7 signifies "No position"
               //because no code was detected. An evaluation that indicates poor quality as the outcome can be due to
               //a misalignment or incorrect orientation, an incorrect measuring distance, or because the code tape has been affixed incorrectly
           END_REGION
       END_REGION

       REGION SICK BARCODE LECTORS
           IF "Control_DB".VTDBarcode_Station[4].Running AND "SICK_Lector_Control_DB_4".Result <> "Control_DB".VTDBarcode_Station[4].Barcode_Old THEN
               "Control_DB".VTD_Sys[4].Inputs."Barcode 1" := "SICK_Lector_Control_DB_4".Result;
               // "Control_DB".VTD_Control.Inputs."Barcode 2'" := SICK_Barcode_DB".Result;
               // "Control_DB".VTDBarcode_Station[4].Barcode_Old := "SICK_Lector_Control_DB_4".Result;
           ELSE
               "Control_DB".VTD_Sys[4].Inputs."Barcode 1" :=
               "Control_DB".VTD_Sys[4].Inputs."Barcode 2" := '';
           END_IF;

       END_REGION

       REGION VFD HARDWARE ID
           //Buffer conveyors 1
           "Settings_DB".LCnv_Sys[4].Cnv_Level[1].Cnv1.G120_Hardware_ID := "C4101~Drive_1~Standard_telegram_20__PZD-2_6";
           "Settings_DB".LCnv_Sys[4].Cnv_Level[2].Cnv1.G120_Hardware_ID := "C4102~Drive_1~Standard_telegram_20__PZD-2_6";
           "Settings_DB".LCnv_Sys[4].Cnv_Level[3].Cnv1.G120_Hardware_ID := "C4103~Drive_1~Standard_telegram_20__PZD-2_6";
           "Settings_DB".LCnv_Sys[4].Cnv_Level[4].Cnv1.G120_Hardware_ID := "C4104~Drive_1~Standard_telegram_20__PZD-2_6";
           "Settings_DB".LCnv_Sys[4].Cnv_Level[5].Cnv1.G120_Hardware_ID := "C4105~Drive_1~Standard_telegram_20__PZD-2_6";
           "Settings_DB".LCnv_Sys[4].Cnv_Level[6].Cnv1.G120_Hardware_ID := "C4106~Drive_1~Standard_telegram_20__PZD-2_6";
           "Settings_DB".LCnv_Sys[4].Cnv_Level[7].Cnv1.G120_Hardware_ID := "C4107~Drive_1~Standard_telegram_20__PZD-2_6";
           "Settings_DB".LCnv_Sys[4].Cnv_Level[8].Cnv1.G120_Hardware_ID := "C4108~Drive_1~Standard_telegram_20__PZD-2_6";

           //Extractor conveyor
           "Settings_DB".ECnv_Sys[4].G120_Hardware_ID := "CVTD_4~Drive_1~Standard_telegram_20__PZD-2_6";

           //VTD
           "Settings_DB".VTD_Sys[4].G120_Hardware_ID := "VTD_4~DO_VECTOR_1~Standard_telegram_20__PZD-2_6";
       END_REGION
   END_REGION

   REGION SYSTEM 5
       REGION EXTRACTOR CONVEYOR
           "Control_DB".ECnv_Sys[5].Inputs.Left := "CVTD5 SENSOR CONVEYOR LEFT (FWD)";
           "Control_DB".ECnv_Sys[5].Inputs.Lpd1 := "CVTD5 SENSOR CONVEYOR LEFT (PALLET DETECT 1)";
           "Control_DB".ECnv_Sys[5].Inputs.Center := "CVTD5 SENSOR CONVEYOR CENTER";
           "Control_DB".ECnv_Sys[5].Inputs.Right := "CVTD5 SENSOR CONVEYOR RIGHT (BWD)";
           "Control_DB".ECnv_Sys[5].Inputs.Rpd1 := "CVTD5 SENSOR CONVEYOR RIGHT (PALLET DETECT 1)";

           "T_OH_Left_5".TOF(IN := "CVTD5 OVERHANG LEFT" OR NOT "Control_DB".VTD_Sys[5].Running,
                             PT := T#200ms);
           "Control_DB".ECnv_Sys[5].Inputs.Overhang_Left := "T_OH_Left_5".Q;
           "I_OH_Right_5".TOF(IN := "CVTD5 OVERHANG RIGHT" OR NOT "Control_DB".VTD_Sys[5].Running,
                             PT := T#200ms);
           "Control_DB".ECnv_Sys[5].Inputs.Overhang_Right := "I_OH_Right_5".Q;

           "Control_DB".ECnv_Sys[5].Inputs.VFD_Status := "CVTD5_StatusWord";
           "Control_DB".ECnv_Sys[5].Inputs.VFD_ActualCurrent := WORD_TO_INT("CVTD5_ActualCurrent");
           "Control_DB".ECnv_Sys[5].Inputs.VFD_Speed_Actual := WORD_TO_INT("CVTD5_ActualSpeed");
           "Control_DB".ECnv_Sys[5].Inputs.VFD_ActualTorque := WORD_TO_INT("CVTD5_ActualTorque");
       END_REGION

       REGION BUFFER CONVEYORS
           REGION LEVEL 1
               //BUFFER CONVEYOR LEVEL 1 - CONVEYOR 1
               "Control_DB".LCnv_Sys[5].Cnv_Level[1].Cnv1.Inputs.Left := NOT "C5101 - SENSOR CNV LEFT (FWD)";
               "Control_DB".LCnv_Sys[5].Cnv_Level[1].Cnv1.Inputs.Lpd1 := NOT "C5101 - SENSOR CNV LEFT (PALLET DETECT 1)";
               "Control_DB".LCnv_Sys[5].Cnv_Level[1].Cnv1.Inputs.Lpd2 := NOT "C5101 - SENSOR CNV LEFT (PALLET DETECT 2)";
               "Control_DB".LCnv_Sys[5].Cnv_Level[1].Cnv1.Inputs.Right := NOT "C5101 - SENSOR CNV RIGHT (BWD)";
               "Control_DB".LCnv_Sys[5].Cnv_Level[1].Cnv1.Inputs.Rpd1 := NOT "C5101 - SENSOR CNV RIGHT (PALLET DETECT 1)";
               "Control_DB".LCnv_Sys[5].Cnv_Level[1].Cnv1.Inputs.Rpd2 := NOT "C5101 - SENSOR CNV RIGHT (PALLET DETECT 2)";
               "Control_DB".LCnv_Sys[5].Cnv_Level[1].Cnv1.Inputs.Sdetect1 := NOT "C5101 - SHUTTLE IN POSITION 1";
               "Control_DB".LCnv_Sys[5].Cnv_Level[1].Cnv1.Inputs.Sdetect2 := NOT "C5101 - SHUTTLE IN POSITION 2";
               "Control_DB".LCnv_Sys[5].Cnv_Level[1].Cnv1.Safety_Stop_Cnrl.Inputs.DP_Extended := "C5101 - SENSOR SAFETY PIN1 UP";
               "Control_DB".LCnv_Sys[5].Cnv_Level[1].Cnv1.Safety_Stop_Cnrl.Inputs.DP_Retracted := "C5101 - SENSOR SAFETY PIN1 DOWN";

               "Control_DB".LCnv_Sys[5].Cnv_Level[1].Cnv1.Inputs.VFD_Status := "C5101_StatusWord";
               "Control_DB".LCnv_Sys[5].Cnv_Level[1].Cnv1.Inputs.VFD_ActualCurrent := WORD_TO_INT("C5101_ActualCurrent");
               "Control_DB".LCnv_Sys[5].Cnv_Level[1].Cnv1.Inputs.VFD_Speed_Actual := WORD_TO_INT("C5101_ActualSpeed");
               "Control_DB".LCnv_Sys[5].Cnv_Level[1].Cnv1.Inputs.VFD_ActualTorque := WORD_TO_INT("C5101_ActualTorque");
           END_REGION

           REGION LEVEL 2
               //BUFFER CONVEYOR LEVEL 2 - CONVEYOR 1
               "Control_DB".LCnv_Sys[5].Cnv_Level[2].Cnv1.Inputs.Left := NOT "C5102 - SENSOR CNV LEFT (FWD)";
               "Control_DB".LCnv_Sys[5].Cnv_Level[2].Cnv1.Inputs.Lpd1 := NOT "C5102 - SENSOR CNV LEFT (PALLET DETECT 1)";
               "Control_DB".LCnv_Sys[5].Cnv_Level[2].Cnv1.Inputs.Lpd2 := NOT "C5102 - SENSOR CNV LEFT (PALLET DETECT 2)";
               "Control_DB".LCnv_Sys[5].Cnv_Level[2].Cnv1.Inputs.Right := NOT "C5102 - SENSOR CNV RIGHT (BWD)";
               "Control_DB".LCnv_Sys[5].Cnv_Level[2].Cnv1.Inputs.Rpd1 := NOT "C5102 - SENSOR CNV RIGHT (PALLET DETECT 1)";
               "Control_DB".LCnv_Sys[5].Cnv_Level[2].Cnv1.Inputs.Rpd2 := NOT "C5102 - SENSOR CNV RIGHT (PALLET DETECT 2)";
               "Control_DB".LCnv_Sys[5].Cnv_Level[2].Cnv1.Inputs.Sdetect1 := NOT "C5102 - SHUTTLE IN POSITION 1";
               "Control_DB".LCnv_Sys[5].Cnv_Level[2].Cnv1.Inputs.Sdetect2 := NOT "C5102 - SHUTTLE IN POSITION 2";
               "Control_DB".LCnv_Sys[5].Cnv_Level[2].Cnv1.Safety_Stop_Cnrl.Inputs.DP_Extended := "C5102 - SENSOR SAFETY PIN1 UP";
               "Control_DB".LCnv_Sys[5].Cnv_Level[2].Cnv1.Safety_Stop_Cnrl.Inputs.DP_Retracted := "C5102 - SENSOR SAFETY PIN1 DOWN";

               "Control_DB".LCnv_Sys[5].Cnv_Level[2].Cnv1.Inputs.VFD_Status := "C5102_StatusWord";
               "Control_DB".LCnv_Sys[5].Cnv_Level[2].Cnv1.Inputs.VFD_ActualCurrent := WORD_TO_INT("C5102_ActualCurrent");
               "Control_DB".LCnv_Sys[5].Cnv_Level[2].Cnv1.Inputs.VFD_Speed_Actual := WORD_TO_INT("C5102_ActualSpeed");
               "Control_DB".LCnv_Sys[5].Cnv_Level[2].Cnv1.Inputs.VFD_ActualTorque := WORD_TO_INT("C5102_ActualTorque");
           END_REGION

           REGION LEVEL 3
               //BUFFER CONVEYOR LEVEL 3 - CONVEYOR 1
               "Control_DB".LCnv_Sys[5].Cnv_Level[3].Cnv1.Inputs.Left := NOT "C5103 - SENSOR CNV LEFT (FWD)";
               "Control_DB".LCnv_Sys[5].Cnv_Level[3].Cnv1.Inputs.Lpd1 := NOT "C5103 - SENSOR CNV LEFT (PALLET DETECT 1)";
               "Control_DB".LCnv_Sys[5].Cnv_Level[3].Cnv1.Inputs.Lpd2 := NOT "C5103 - SENSOR CNV LEFT (PALLET DETECT 2)";
               "Control_DB".LCnv_Sys[5].Cnv_Level[3].Cnv1.Inputs.Right := NOT "C5103 - SENSOR CNV RIGHT (BWD)";
               "Control_DB".LCnv_Sys[5].Cnv_Level[3].Cnv1.Inputs.Rpd1 := NOT "C5103 - SENSOR CNV RIGHT (PALLET DETECT 1)";
               "Control_DB".LCnv_Sys[5].Cnv_Level[3].Cnv1.Inputs.Rpd2 := NOT "C5103 - SENSOR CNV RIGHT (PALLET DETECT 2)";
               "Control_DB".LCnv_Sys[5].Cnv_Level[3].Cnv1.Inputs.Sdetect1 := NOT "C5103 - SHUTTLE IN POSITION 1";
               "Control_DB".LCnv_Sys[5].Cnv_Level[3].Cnv1.Inputs.Sdetect2 := NOT "C5103 - SHUTTLE IN POSITION 2";
               "Control_DB".LCnv_Sys[5].Cnv_Level[3].Cnv1.Safety_Stop_Cnrl.Inputs.DP_Extended := "C5103 - SENSOR SAFETY PIN1 UP";
               "Control_DB".LCnv_Sys[5].Cnv_Level[3].Cnv1.Safety_Stop_Cnrl.Inputs.DP_Retracted := "C5103 - SENSOR SAFETY PIN1 DOWN";

               "Control_DB".LCnv_Sys[5].Cnv_Level[3].Cnv1.Inputs.VFD_Status := "C5103_StatusWord";
               "Control_DB".LCnv_Sys[5].Cnv_Level[3].Cnv1.Inputs.VFD_ActualCurrent := WORD_TO_INT("C5103_ActualCurrent");
               "Control_DB".LCnv_Sys[5].Cnv_Level[3].Cnv1.Inputs.VFD_Speed_Actual := WORD_TO_INT("C5103_ActualSpeed");
               "Control_DB".LCnv_Sys[5].Cnv_Level[3].Cnv1.Inputs.VFD_ActualTorque := WORD_TO_INT("C5103_ActualTorque");
           END_REGION

           REGION LEVEL 4
               //BUFFER CONVEYOR LEVEL 4 - CONVEYOR 1
               "Control_DB".LCnv_Sys[5].Cnv_Level[4].Cnv1.Inputs.Left := NOT "C5104 - SENSOR CNV LEFT (FWD)";
               "Control_DB".LCnv_Sys[5].Cnv_Level[4].Cnv1.Inputs.Lpd1 := NOT "C5104 - SENSOR CNV LEFT (PALLET DETECT 1)";
               "Control_DB".LCnv_Sys[5].Cnv_Level[4].Cnv1.Inputs.Lpd2 := NOT "C5104 - SENSOR CNV LEFT (PALLET DETECT 2)";
               "Control_DB".LCnv_Sys[5].Cnv_Level[4].Cnv1.Inputs.Right := NOT "C5104 - SENSOR CNV RIGHT (BWD)";
               "Control_DB".LCnv_Sys[5].Cnv_Level[4].Cnv1.Inputs.Rpd1 := NOT "C5104 - SENSOR CNV RIGHT (PALLET DETECT 1)";
               "Control_DB".LCnv_Sys[5].Cnv_Level[4].Cnv1.Inputs.Rpd2 := NOT "C5104 - SENSOR CNV RIGHT (PALLET DETECT 2)";
               "Control_DB".LCnv_Sys[5].Cnv_Level[4].Cnv1.Inputs.Sdetect1 := NOT "C5104 - SHUTTLE IN POSITION 1";
               "Control_DB".LCnv_Sys[5].Cnv_Level[4].Cnv1.Inputs.Sdetect2 := NOT "C5104 - SHUTTLE IN POSITION 2";
               "Control_DB".LCnv_Sys[5].Cnv_Level[4].Cnv1.Safety_Stop_Cnrl.Inputs.DP_Extended := "C5104 - SENSOR SAFETY PIN1 UP";
               "Control_DB".LCnv_Sys[5].Cnv_Level[4].Cnv1.Safety_Stop_Cnrl.Inputs.DP_Retracted := "C5104 - SENSOR SAFETY PIN1 DOWN";

               "Control_DB".LCnv_Sys[5].Cnv_Level[4].Cnv1.Inputs.VFD_Status := "C5104_StatusWord";
               "Control_DB".LCnv_Sys[5].Cnv_Level[4].Cnv1.Inputs.VFD_ActualCurrent := WORD_TO_INT("C5104_ActualCurrent");
               "Control_DB".LCnv_Sys[5].Cnv_Level[4].Cnv1.Inputs.VFD_Speed_Actual := WORD_TO_INT("C5104_ActualSpeed");
               "Control_DB".LCnv_Sys[5].Cnv_Level[4].Cnv1.Inputs.VFD_ActualTorque := WORD_TO_INT("C5104_ActualTorque");
           END_REGION

           REGION LEVEL 5
               //BUFFER CONVEYOR LEVEL 5 - CONVEYOR 1
               "Control_DB".LCnv_Sys[5].Cnv_Level[5].Cnv1.Inputs.Left := NOT "C5105 - SENSOR CNV LEFT (FWD)";
               "Control_DB".LCnv_Sys[5].Cnv_Level[5].Cnv1.Inputs.Lpd1 := NOT "C5105 - SENSOR CNV LEFT (PALLET DETECT 1)";
               "Control_DB".LCnv_Sys[5].Cnv_Level[5].Cnv1.Inputs.Lpd2 := NOT "C5105 - SENSOR CNV LEFT (PALLET DETECT 2)";
               "Control_DB".LCnv_Sys[5].Cnv_Level[5].Cnv1.Inputs.Right := NOT "C5105 - SENSOR CNV RIGHT (BWD)";
               "Control_DB".LCnv_Sys[5].Cnv_Level[5].Cnv1.Inputs.Rpd1 := NOT "C5105 - SENSOR CNV RIGHT (PALLET DETECT 1)";
               "Control_DB".LCnv_Sys[5].Cnv_Level[5].Cnv1.Inputs.Rpd2 := NOT "C5105 - SENSOR CNV RIGHT (PALLET DETECT 2)";
               "Control_DB".LCnv_Sys[5].Cnv_Level[5].Cnv1.Inputs.Sdetect1 := NOT "C5105 - SHUTTLE IN POSITION 1";
               "Control_DB".LCnv_Sys[5].Cnv_Level[5].Cnv1.Inputs.Sdetect2 := NOT "C5105 - SHUTTLE IN POSITION 2";
               "Control_DB".LCnv_Sys[5].Cnv_Level[5].Cnv1.Safety_Stop_Cnrl.Inputs.DP_Extended := "C5105 - SENSOR SAFETY PIN1 UP";
               "Control_DB".LCnv_Sys[5].Cnv_Level[5].Cnv1.Safety_Stop_Cnrl.Inputs.DP_Retracted := "C5105 - SENSOR SAFETY PIN1 DOWN";

               "Control_DB".LCnv_Sys[5].Cnv_Level[5].Cnv1.Inputs.VFD_Status := "C5105_StatusWord";
               "Control_DB".LCnv_Sys[5].Cnv_Level[5].Cnv1.Inputs.VFD_ActualCurrent := WORD_TO_INT("C5105_ActualCurrent");
               "Control_DB".LCnv_Sys[5].Cnv_Level[5].Cnv1.Inputs.VFD_Speed_Actual := WORD_TO_INT("C5105_ActualSpeed");
               "Control_DB".LCnv_Sys[5].Cnv_Level[5].Cnv1.Inputs.VFD_ActualTorque := WORD_TO_INT("C5105_ActualTorque");
           END_REGION

           REGION LEVEL 6
               //BUFFER CONVEYOR LEVEL 6 - CONVEYOR 1
               "Control_DB".LCnv_Sys[5].Cnv_Level[6].Cnv1.Inputs.Left := NOT "C5106 - SENSOR CNV LEFT (FWD)";
               "Control_DB".LCnv_Sys[5].Cnv_Level[6].Cnv1.Inputs.Lpd1 := NOT "C5106 - SENSOR CNV LEFT (PALLET DETECT 1)";
               "Control_DB".LCnv_Sys[5].Cnv_Level[6].Cnv1.Inputs.Lpd2 := NOT "C5106 - SENSOR CNV LEFT (PALLET DETECT 2)";
               "Control_DB".LCnv_Sys[5].Cnv_Level[6].Cnv1.Inputs.Right := NOT "C5106 - SENSOR CNV RIGHT (BWD)";
               "Control_DB".LCnv_Sys[5].Cnv_Level[6].Cnv1.Inputs.Rpd1 := NOT "C5106 - SENSOR CNV RIGHT (PALLET DETECT 1)";
               "Control_DB".LCnv_Sys[5].Cnv_Level[6].Cnv1.Inputs.Rpd2 := NOT "C5106 - SENSOR CNV RIGHT (PALLET DETECT 2)";
               "Control_DB".LCnv_Sys[5].Cnv_Level[6].Cnv1.Inputs.Sdetect1 := NOT "C5106 - SHUTTLE IN POSITION 1";
               "Control_DB".LCnv_Sys[5].Cnv_Level[6].Cnv1.Inputs.Sdetect2 := NOT "C5106 - SHUTTLE IN POSITION 2";
               "Control_DB".LCnv_Sys[5].Cnv_Level[6].Cnv1.Safety_Stop_Cnrl.Inputs.DP_Extended := "C5106 - SENSOR SAFETY PIN1 UP";
               "Control_DB".LCnv_Sys[5].Cnv_Level[6].Cnv1.Safety_Stop_Cnrl.Inputs.DP_Retracted := "C5106 - SENSOR SAFETY PIN1 DOWN";

               "Control_DB".LCnv_Sys[5].Cnv_Level[6].Cnv1.Inputs.VFD_Status := "C5106_StatusWord";
               "Control_DB".LCnv_Sys[5].Cnv_Level[6].Cnv1.Inputs.VFD_ActualCurrent := WORD_TO_INT("C5106_ActualCurrent");
               "Control_DB".LCnv_Sys[5].Cnv_Level[6].Cnv1.Inputs.VFD_Speed_Actual := WORD_TO_INT("C5106_ActualSpeed");
               "Control_DB".LCnv_Sys[5].Cnv_Level[6].Cnv1.Inputs.VFD_ActualTorque := WORD_TO_INT("C5106_ActualTorque");
           END_REGION

           REGION LEVEL 7
               //BUFFER CONVEYOR LEVEL 7 - CONVEYOR 1
               "Control_DB".LCnv_Sys[5].Cnv_Level[7].Cnv1.Inputs.Left := NOT "C5107 - SENSOR CNV LEFT (FWD)";
               "Control_DB".LCnv_Sys[5].Cnv_Level[7].Cnv1.Inputs.Lpd1 := NOT "C5107 - SENSOR CNV LEFT (PALLET DETECT 1)";
               "Control_DB".LCnv_Sys[5].Cnv_Level[7].Cnv1.Inputs.Lpd2 := NOT "C5107 - SENSOR CNV LEFT (PALLET DETECT 2)";
               "Control_DB".LCnv_Sys[5].Cnv_Level[7].Cnv1.Inputs.Right := NOT "C5107 - SENSOR CNV RIGHT (BWD)";
               "Control_DB".LCnv_Sys[5].Cnv_Level[7].Cnv1.Inputs.Rpd1 := NOT "C5107 - SENSOR CNV RIGHT (PALLET DETECT 1)";
               "Control_DB".LCnv_Sys[5].Cnv_Level[7].Cnv1.Inputs.Rpd2 := NOT "C5107 - SENSOR CNV RIGHT (PALLET DETECT 2)";
               "Control_DB".LCnv_Sys[5].Cnv_Level[7].Cnv1.Inputs.Sdetect1 := NOT "C5107 - SHUTTLE IN POSITION 1";
               "Control_DB".LCnv_Sys[5].Cnv_Level[7].Cnv1.Inputs.Sdetect2 := NOT "C5107 - SHUTTLE IN POSITION 2";
               "Control_DB".LCnv_Sys[5].Cnv_Level[7].Cnv1.Safety_Stop_Cnrl.Inputs.DP_Extended := "C5107 - SENSOR SAFETY PIN1 UP";
               "Control_DB".LCnv_Sys[5].Cnv_Level[7].Cnv1.Safety_Stop_Cnrl.Inputs.DP_Retracted := "C5107 - SENSOR SAFETY PIN1 DOWN";

               "Control_DB".LCnv_Sys[5].Cnv_Level[7].Cnv1.Inputs.VFD_Status := "C5107_StatusWord";
               "Control_DB".LCnv_Sys[5].Cnv_Level[7].Cnv1.Inputs.VFD_ActualCurrent := WORD_TO_INT("C5107_ActualCurrent");
               "Control_DB".LCnv_Sys[5].Cnv_Level[7].Cnv1.Inputs.VFD_Speed_Actual := WORD_TO_INT("C5107_ActualSpeed");
               "Control_DB".LCnv_Sys[5].Cnv_Level[7].Cnv1.Inputs.VFD_ActualTorque := WORD_TO_INT("C5107_ActualTorque");
           END_REGION

           REGION LEVEL 8
               //BUFFER CONVEYOR LEVEL 8 - CONVEYOR 1
               "Control_DB".LCnv_Sys[5].Cnv_Level[8].Cnv1.Inputs.Left := NOT "C5108 - SENSOR CNV LEFT (FWD)";
               "Control_DB".LCnv_Sys[5].Cnv_Level[8].Cnv1.Inputs.Lpd1 := NOT "C5108 - SENSOR CNV LEFT (PALLET DETECT 1)";
               "Control_DB".LCnv_Sys[5].Cnv_Level[8].Cnv1.Inputs.Lpd2 := NOT "C5108 - SENSOR CNV LEFT (PALLET DETECT 2)";
               "Control_DB".LCnv_Sys[5].Cnv_Level[8].Cnv1.Inputs.Right := NOT "C5108 - SENSOR CNV RIGHT (BWD)";
               "Control_DB".LCnv_Sys[5].Cnv_Level[8].Cnv1.Inputs.Rpd1 := NOT "C5108 - SENSOR CNV RIGHT (PALLET DETECT 1)";
               "Control_DB".LCnv_Sys[5].Cnv_Level[8].Cnv1.Inputs.Rpd2 := NOT "C5108 - SENSOR CNV RIGHT (PALLET DETECT 2)";
               "Control_DB".LCnv_Sys[5].Cnv_Level[8].Cnv1.Inputs.Sdetect1 := NOT "C5108 - SHUTTLE IN POSITION 1";
               "Control_DB".LCnv_Sys[5].Cnv_Level[8].Cnv1.Inputs.Sdetect2 := NOT "C5108 - SHUTTLE IN POSITION 2";
               "Control_DB".LCnv_Sys[5].Cnv_Level[8].Cnv1.Safety_Stop_Cnrl.Inputs.DP_Extended := "C5108 - SENSOR SAFETY PIN1 UP";
               "Control_DB".LCnv_Sys[5].Cnv_Level[8].Cnv1.Safety_Stop_Cnrl.Inputs.DP_Retracted := "C5108 - SENSOR SAFETY PIN1 DOWN";

               "Control_DB".LCnv_Sys[5].Cnv_Level[8].Cnv1.Inputs.VFD_Status := "C5108_StatusWord";
               "Control_DB".LCnv_Sys[5].Cnv_Level[8].Cnv1.Inputs.VFD_ActualCurrent := WORD_TO_INT("C5108_ActualCurrent");
               "Control_DB".LCnv_Sys[5].Cnv_Level[8].Cnv1.Inputs.VFD_Speed_Actual := WORD_TO_INT("C5108_ActualSpeed");
               "Control_DB".LCnv_Sys[5].Cnv_Level[8].Cnv1.Inputs.VFD_ActualTorque := WORD_TO_INT("C5108_ActualTorque");
           END_REGION
       END_REGION

       REGION VTD
           "Control_DB".VTD_Sys[5].Inputs.Upper_Overtravel := "OVERTRAVEL UPPER LIMIT - CH1(5)";
           "Control_DB".VTD_Sys[5].Inputs.Upper_limit := "VTD5 UPPER LIMIT";
           "Control_DB".VTD_Sys[5].Inputs.Ultimate_SlowDown := "VTD5 ULTIMATE SLOWDOWN";
           "Control_DB".VTD_Sys[5].Inputs.Ultimate_Creep := "VTD5 ULTIMATE CREEP";
           "Control_DB".VTD_Sys[5].Inputs.Lower_Limit := "VTD5 LOWER LIMIT";
           "Control_DB".VTD_Sys[5].Inputs.Lower_Overtravel := "OVERTRAVEL LOWER LIMIT - CH1(5)";
           "Control_DB".VTD_Sys[5].Inputs.Level_Detect1 := "VTD5 LEVEL DETECT 1";
           "Control_DB".VTD_Sys[5].Inputs.Level_Detect2 := "VTD5 LEVEL DETECT 2";
           "Control_DB".VTD_Sys[5].Inputs.DP1_Extended := "VTD5 DOCKING PINS 1 EXTENDED";
           "Control_DB".VTD_Sys[5].Inputs.DP2_Extended := "VTD5 DOCKING PINS 2 EXTENDED";
           "Control_DB".VTD_Sys[5].Inputs.DP1_Retracted := "VTD5 DOCKING PINS 1 RETRACTED";
           "Control_DB".VTD_Sys[5].Inputs.DP2_Retracted := "VTD5 DOCKING PINS 2 RETRACTED";
           "Control_DB".VTD_Sys[5].Inputs.Chain_Slack_1 := NOT "Remote_Panel_DB_5".Chain_Slack_1_Filtered;
           "Control_DB".VTD_Sys[5].Inputs.Chain_Slack_2 := NOT "Remote_Panel_DB_5".Chain_Slack_2_Filtered;
           "Control_DB".VTD_Sys[5].Inputs.Chain_Slack_3 := NOT "Remote_Panel_DB_5".Chain_Slack_3_Filtered;
           "Control_DB".VTD_Sys[5].Inputs.Chain_Slack_4 := NOT "Remote_Panel_DB_5".Chain_Slack_4_Filtered;
           "Control_DB".VTD_Sys[5].Inputs.PushToEnter := "VTD5 PUSH TO ENTER VTD ZONE";
           "Control_DB".VTD_Sys[5].Inputs.PushToExit := "VTD5 PUSH TO EXIT VTD ZONE";
           "Control_DB".VTD_Sys[5].Inputs.VFD_Status := "VTD5_StatusWord";
           "Control_DB".VTD_Sys[5].Inputs.VFD_ActualCurrent := REAL_TO_INT(("VTD5_ActualCurrent" / 10) / 72.5);
           "Control_DB".VTD_Sys[5].Inputs.VFD_Speed_Actual := "VTD5_ActualSpeed";
           "Control_DB".VTD_Sys[5].Inputs.VFD_ActualTorque := WORD_TO_INT("VTD5_ActualTorque");

       END_REGION

       REGION ABSOLUTE ENCODER
           REGION DOCUMENTATION
               //STATUS---------------------------------------------------------------------------------------------------------------------
               //
               //Encoder state word 2 - INPUT WORD 1
               //
               // 15 … 12 Encoder’s Sign-OF-Life (NOT relevant)
               // 11, 10 Reserved
               // 9 Control requested 0 = No control BY the PLC requested 1 = Control BY the PLC requested
               // 8 … 0 Reserved

               //Sensor 1 state word - INPUT WORD 2
               //
               // 15 Encoder error Description 0 = No error 1 = Error The error code is output in G1_XIST2.
               // 14 Park mode activated 0 = Normal operation 1 = Park mode activated Feedback based on G1_STW bit 14: No output OF position data G1_XIST1 AND G1_XIST2
               // 13 Transmission OF absolute position value 0 = No transmission 1 = Position value is output in G1_XIST2
               // 12 Status OF the Preset function (set/shift OF home position executed) 0 = No Preset function active 1 = Preset function is run Feedback based on G1_STW bit 12:  
               // 11 Requirement OF error acknowledgement detected New position value is output in G1_XIST1 AND G1_XIST2. On conclusion OF the Preset function the bit is set TO 0. 0 = No RETURN acknowledgement OF Encoder error 1 = Requirement OF error acknowledgement detected Reaction TO bit 15 in the sensor control word 1 G1_STW is acknowledged (see Table 14)
               // 10 Reserved
               // 9 … 0 NOT supported

               //Position 1 - INPUT WORD 3 AND 4
               // "AE_Position_1_Scaled" := (*SCALE_X(MIN := "Settings_DB".VTD_Settings.VTD_Min_Height,
               //                                   VALUE := *)NORM_X(MIN := 0,
               //                                                   VALUE := (SHL(IN:="AE_Position_1", N:=2) * 0.00228881) (*- "AE_Offset"*),
               //                                                   MAX := 1073741824)(*,
               //                                   MAX := "Settings_DB".VTD_Settings.VTD_Max_Heigh)*);
               // "mm_per_pulse" := 401,5584 / 262144;
               // 
               //CONTROL---------------------------------------------------------------------------------------------------------------------
               //
               //Encoder control word 2 - OUTPUT WORD 1
               //
               // 15 … 12 Master’s Sign-OF-Life (NOT relevant)
               // 10 control BY PLC 0 = No control BY the PLC 1 = Control BY the PLC Enables the PLC BY using control words TO activate / deactivate encoder functions
               // 7 Fault acknowledge Error-buffer handling NOT supported
               // 11, 9, 8, 6 … 0 Reserved
               // "AE_Control_Word_1".%X10 := "AE_PLC_Control";
               // 
               //Sensor 1 control word - OUTPUT WORD 2-------------------------------------------------------------------------------------------
               //
               // 15 Acknowledging a sensor error Description 0 = Encoder error message NOT acknowledged BY PLC 1 = Encoder error message acknowledged BY the PLC
               // 14 Activate park mode 0 = Normal operation 1 = Activate park mode
               // 13 Request FOR the absolute position value 0 = No request 1 = Request BY the master Results in the cyclic output OF the position values in G1_XIST2
               // 12 Activate preset value (see note below) Defines that a configured preset value is used (see section 3.5 on page 24) 0 = Preset value is NOT activated 1 = Preset value is activated
               // 11 Preset mode Defines how a configured preset value is used 0 = Preset value is used as a new absolute value 1 = Preset value is added TO the previous value
               // 10 … 0 Reserved
               // "AE_Control_Word_2".%X15 := "VTD_Reset_HMI_Tags";
               // "AE_Control_Word_2".%X14 := "AE_Activate_ParkMode";
               // "AE_Control_Word_2".%X13 := "AE_Request_ABS_Value";
               // "AE_Control_Word_2".%X12 := "AE_Activate_Preset_Value";
               // "AE_Control_Word_2".%X11 := "AE_Preset_Mode";
           END_REGION

           //STATUS---------------------------------------------------------------------------------------------------------------------
           "Control_DB".VTD_Sys[5].Inputs.AE_Status_2 := "AE_Status_2(5)";
           //Position 1 - INPUT WORD 3 AND 4
           "Control_DB".VTD_Sys[5].Inputs.AE_Position_1 := REAL_TO_DINT((((1073741823 - (*reverse the direction*)
    (SHR(IN := "AE_Position_1(5)", N := 2))) - 31381317) * 0.0015318237304688 (*Mechanical relationship*) - 1805195)(*Offset*));

   // Position 2 - INPUT WORD 5 AND 6
           "Control_DB".VTD_Sys[5].Inputs.AE_Position_2 := SHR(IN := "AE_Position_2(5)", N := 2);

           //Speed A - INPUT WORD 7
           "Control_DB".VTD_Sys[5].Inputs.AE_Speed := "AE_Speed(5)";
       END_REGION

       REGION LINEAR ENCODER
           "Control_DB".VTD_Sys[5].Inputs.LE_Position := "LE_X_Unsafe_Position(5)" / 10;
           "Control_DB".VTD_Sys[5].Inputs.LE_Speed := "LE_Speed(5)" * 100;
           "Control_DB".VTD_Sys[5].Inputs.LE_Status := "LE_Status(5)";
           "Control_DB".VTD_Sys[5].Inputs.LE_Warnings := "LE_Warnings(5)";
           REGION DOCUMENTATION
               //STATUS 
               //
               // 0 ERR - Error message (Error code in XP00– XP15); remaining bits = 0, see Error Codes
               // 1 NP - No position information/OUT (XP = 0, YP = 0, SP = 0)
               // 2 WRN - Warnings present, see Warning Module
               // 3 EV - Event present
               // 4 posdetected - Valid position information available

               //WARNINGS
               //
               // 0 WRN01 A code with non-PXV content was found.
               // 1 WRN02 the read head is too close TO the Data Matrix code tape.
               // 2 WRN03 the read head is too far from the Data Matrix code tape.
               // 3 WRN04 Y position too large. The sensor is just before OUT.
               // 4 WRN05 Y position is too small. The sensor is just before OUT.
               // 5 WRN06 the read head is rotated OR tilted in relation TO the Data Matrix code tape.
               // 6 WRN07 Low level OF code contrast.
               // 7 WRN08 Repair tape detected.
               // 8 WRN09 Temperature too high.
               // 9...15 Reserved

               //QUALITY GRADE
               //
               //The quality grades enable constant monitoring of the code tape and the camera along the entire
               //traverse distance. This enables you to detect and act upon potential damage or contamination
               //of the code tape and camera at the earliest stage possible during commissioning and normal
               //operation. As a result, this maximizes the overall functional reliability of your plant, and
               //it means you are able to immediately localize the issue in the case of a fault. Evaluations
               //are made using a scale of 1 to 6. The value 1 is the best possible read quality. A value greater
               //than 3 or worse requires the camera and its path to be inspected. The value 7 signifies "No position"
               //because no code was detected. An evaluation that indicates poor quality as the outcome can be due to
               //a misalignment or incorrect orientation, an incorrect measuring distance, or because the code tape has been affixed incorrectly
           END_REGION
       END_REGION

       REGION SICK BARCODE LECTORS
           IF "Control_DB".VTDBarcode_Station[5].Running AND "SICK_Lector_Control_DB_5".Result <> "Control_DB".VTDBarcode_Station[5].Barcode_Old THEN
               "Control_DB".VTD_Sys[5].Inputs."Barcode 1" := "SICK_Lector_Control_DB_5".Result;
               // "Control_DB".VTD_Control.Inputs."Barcode 2'" := SICK_Barcode_DB".Result;
               // "Control_DB".VTDBarcode_Station[5].Barcode_Old := "SICK_Lector_Control_DB_5".Result;
           ELSE
               "Control_DB".VTD_Sys[5].Inputs."Barcode 1" :=
               "Control_DB".VTD_Sys[5].Inputs."Barcode 2" := '';
           END_IF;

       END_REGION

       REGION VFD HARDWARE ID
           //Buffer conveyors 1
           "Settings_DB".LCnv_Sys[5].Cnv_Level[1].Cnv1.G120_Hardware_ID := "C5101~Drive_1~Standard_telegram_20__PZD-2_6";
           "Settings_DB".LCnv_Sys[5].Cnv_Level[2].Cnv1.G120_Hardware_ID := "C5102~Drive_1~Standard_telegram_20__PZD-2_6";
           "Settings_DB".LCnv_Sys[5].Cnv_Level[3].Cnv1.G120_Hardware_ID := "C5103~Drive_1~Standard_telegram_20__PZD-2_6";
           "Settings_DB".LCnv_Sys[5].Cnv_Level[4].Cnv1.G120_Hardware_ID := "C5104~Drive_1~Standard_telegram_20__PZD-2_6";
           "Settings_DB".LCnv_Sys[5].Cnv_Level[5].Cnv1.G120_Hardware_ID := "C5105~Drive_1~Standard_telegram_20__PZD-2_6";
           "Settings_DB".LCnv_Sys[5].Cnv_Level[6].Cnv1.G120_Hardware_ID := "C5106~Drive_1~Standard_telegram_20__PZD-2_6";
           "Settings_DB".LCnv_Sys[5].Cnv_Level[7].Cnv1.G120_Hardware_ID := "C5107~Drive_1~Standard_telegram_20__PZD-2_6";
           "Settings_DB".LCnv_Sys[5].Cnv_Level[8].Cnv1.G120_Hardware_ID := "C5108~Drive_1~Standard_telegram_20__PZD-2_6";

           //Extractor conveyor
           "Settings_DB".ECnv_Sys[5].G120_Hardware_ID := "CVTD_5~Drive_1~Standard_telegram_20__PZD-2_6";

           //VTD
           "Settings_DB".VTD_Sys[5].G120_Hardware_ID := "VTD_5~DO_VECTOR_1~Standard_telegram_20__PZD-2_6";
       END_REGION
   END_REGION

   REGION LEVEL KEYS
       // System 1
       "HMI_DB".Rem_Loc_Keys[1].Level[1] := "KEY REMOTE/LOCAL L1 - CH1(1)";
       "HMI_DB".Rem_Loc_Keys[1].Level[2] := "KEY REMOTE/LOCAL L2 - CH1(1)";
       "HMI_DB".Rem_Loc_Keys[1].Level[3] := "KEY REMOTE/LOCAL L3 - CH1(1)";
       "HMI_DB".Rem_Loc_Keys[1].Level[4] := "KEY REMOTE/LOCAL L4 - CH1(1)";
       "HMI_DB".Rem_Loc_Keys[1].Level[5] := "KEY REMOTE/LOCAL L5 - CH1(1)";
       "HMI_DB".Rem_Loc_Keys[1].Level[6] := "KEY REMOTE/LOCAL L6 - CH1(1)";
       "HMI_DB".Rem_Loc_Keys[1].Level[7] := "KEY REMOTE/LOCAL L7 - CH1(1)";
       "HMI_DB".Rem_Loc_Keys[1].Level[8] := "KEY REMOTE/LOCAL L8 - CH1(1)";

       // System 2
       "HMI_DB".Rem_Loc_Keys[2].Level[1] := "KEY REMOTE/LOCAL L1 - CH1(2)";
       "HMI_DB".Rem_Loc_Keys[2].Level[2] := "KEY REMOTE/LOCAL L2 - CH1(2)";
       "HMI_DB".Rem_Loc_Keys[2].Level[3] := "KEY REMOTE/LOCAL L3 - CH1(2)";
       "HMI_DB".Rem_Loc_Keys[2].Level[4] := "KEY REMOTE/LOCAL L4 - CH1(2)";
       "HMI_DB".Rem_Loc_Keys[2].Level[5] := "KEY REMOTE/LOCAL L5 - CH1(2)";
       "HMI_DB".Rem_Loc_Keys[2].Level[6] := "KEY REMOTE/LOCAL L6 - CH1(2)";
       "HMI_DB".Rem_Loc_Keys[2].Level[7] := "KEY REMOTE/LOCAL L7 - CH1(2)";
       "HMI_DB".Rem_Loc_Keys[2].Level[8] := "KEY REMOTE/LOCAL L8 - CH1(2)";

       // System 3
       "HMI_DB".Rem_Loc_Keys[3].Level[1] := "KEY REMOTE/LOCAL L1 - CH1(3)";
       "HMI_DB".Rem_Loc_Keys[3].Level[2] := "KEY REMOTE/LOCAL L2 - CH1(3)";
       "HMI_DB".Rem_Loc_Keys[3].Level[3] := "KEY REMOTE/LOCAL L3 - CH1(3)";
       "HMI_DB".Rem_Loc_Keys[3].Level[4] := "KEY REMOTE/LOCAL L4 - CH1(3)";
       "HMI_DB".Rem_Loc_Keys[3].Level[5] := "KEY REMOTE/LOCAL L5 - CH1(3)";
       "HMI_DB".Rem_Loc_Keys[3].Level[6] := "KEY REMOTE/LOCAL L6 - CH1(3)";
       "HMI_DB".Rem_Loc_Keys[3].Level[7] := "KEY REMOTE/LOCAL L7 - CH1(3)";
       "HMI_DB".Rem_Loc_Keys[3].Level[8] := "KEY REMOTE/LOCAL L8 - CH1(3)";

       // System 4
       "HMI_DB".Rem_Loc_Keys[4].Level[1] := "KEY REMOTE/LOCAL L1 - CH1(4)";
       "HMI_DB".Rem_Loc_Keys[4].Level[2] := "KEY REMOTE/LOCAL L2 - CH1(4)";
       "HMI_DB".Rem_Loc_Keys[4].Level[3] := "KEY REMOTE/LOCAL L3 - CH1(4)";
       "HMI_DB".Rem_Loc_Keys[4].Level[4] := "KEY REMOTE/LOCAL L4 - CH1(4)";
       "HMI_DB".Rem_Loc_Keys[4].Level[5] := "KEY REMOTE/LOCAL L5 - CH1(4)";
       "HMI_DB".Rem_Loc_Keys[4].Level[6] := "KEY REMOTE/LOCAL L6 - CH1(4)";
       "HMI_DB".Rem_Loc_Keys[4].Level[7] := "KEY REMOTE/LOCAL L7 - CH1(4)";
       "HMI_DB".Rem_Loc_Keys[4].Level[8] := "KEY REMOTE/LOCAL L8 - CH1(4)";

       // System 5
       "HMI_DB".Rem_Loc_Keys[5].Level[1] := "KEY REMOTE/LOCAL L1 - CH1(5)";
       "HMI_DB".Rem_Loc_Keys[5].Level[2] := "KEY REMOTE/LOCAL L2 - CH1(5)";
       "HMI_DB".Rem_Loc_Keys[5].Level[3] := "KEY REMOTE/LOCAL L3 - CH1(5)";
       "HMI_DB".Rem_Loc_Keys[5].Level[4] := "KEY REMOTE/LOCAL L4 - CH1(5)";
       "HMI_DB".Rem_Loc_Keys[5].Level[5] := "KEY REMOTE/LOCAL L5 - CH1(5)";
       "HMI_DB".Rem_Loc_Keys[5].Level[6] := "KEY REMOTE/LOCAL L6 - CH1(5)";
       "HMI_DB".Rem_Loc_Keys[5].Level[7] := "KEY REMOTE/LOCAL L7 - CH1(5)";
       "HMI_DB".Rem_Loc_Keys[5].Level[8] := "KEY REMOTE/LOCAL L8 - CH1(5)";
   END_REGION;
END_FUNCTION

FUNCTION_BLOCK "MQTT_Handler_FB"   // FB2, SCL
{ S7_Optimized_Access := 'TRUE' }
VERSION : 0.1
// stored: AutoNumber true, IsIECCheckEnabled false, IsRetainMemResEnabled false, MemoryReserve 100, SetENOAutomatically false, UDAEnableTagReadback false
   VAR_INPUT
      Enable : Bool := True;
   END_VAR
   VAR_IN_OUT
      LMQTT_DB : "LMQTT_DB_UDT";
   END_VAR
   VAR
      MQTT_Setup : Bool;
      MQTT_Topic : WString;
      Publish_Msg_Payload : Array[1..128] of Byte;
      Received_Topic : WString;
      Received_Msg_Payload : Array[0..1024] of Byte;
      i : UInt;
      j : UInt;
      Subscribe : Bool;
      Unsubscribe : Bool;
      Received_Msg_Status : USInt;
      Received_Msg_Length : UDInt;
      Busy : Bool;
      Valid : Bool;
      Done : Bool;
      Error : Bool;
      Status : Word;
      Diagnostics { S7_SetPoint := 'True'} : "typeDiagnostics";
      JSON_Tree : Array[1..18] of "LStream_typeElement";
      Shuttle_No : UInt;
      sSubTopic : Array[1..24] of String;
      bSubscribed : Bool;
      SubscribeState : Int;
      SubscribeIndex : Int := 1;
      SubscribeCount : UInt := 1;
      SubscribeTopicList : Array[1..30] of String;
      sPayloadRcv : String;
      sPayloadRcv_1 : String;
      sPayloadRcv_2 : String;
      sPayloadRcv_3 : String;
      sPayloadRcv_4 : String;
      sPayloadRcv_5 : String;
      MQTT_AutoReset : UInt;
      Enable_AutoReset : Bool;
      T_AutoReset { S7_SetPoint := 'True'} : TON_TIME;
   END_VAR
   VAR_TEMP
      iIndex : UInt;
      sIndexStr : String;
      k : UInt;
      test : DWord;
      Y : UInt;
   END_VAR
BEGIN
   (*
   TODO
   1. Add timeout on subscribe event
   2. Add cyclic checks for all the different errors in the status word

   Status word values:
   16#0000 Last job (publish/subscribe/unsubscribe) successfully executed
   16#7000 Block is idle/client not connected
   16#7001 First call after "enable" = TRUE
   16#7002 Block processes job
   16#7003 Establishing connection to MQTT broker
   16#7004 MQTT client connected and ready for job
   16#7005 Ping is sent to the broker
   16#7006 Publish job is executed
   16#7008 Subscribe job is executed
   16#7010 Unsubscribe job is executed
   *)

   IF "FirstScan" THEN
       "MQTT_Enable" := TRUE;
   END_IF;

   #LMQTT_DB.connParam := "Settings_DB".Shuttle_MQTT.MQTT_Con_Params;
   #LMQTT_DB.clientIdentifier := "Settings_DB".Shuttle_MQTT.Client_ID;
   #LMQTT_DB.username := "Settings_DB".Shuttle_MQTT.Username;
   #LMQTT_DB.password := "Settings_DB".Shuttle_MQTT.Password;
   #LMQTT_DB.willtopic := "Settings_DB".Shuttle_MQTT.Will_Topic;
   #LMQTT_DB.willMsgPayload := "Settings_DB".Shuttle_MQTT.Will_Msg_Payload;
   #LMQTT_DB.willMsgLen := 0;
   #LMQTT_DB.willMsgPayload := #Publish_Msg_Payload;
   #Received_Topic := #LMQTT_DB.receivedTopic;
   #Received_Msg_Payload := #LMQTT_DB.receivedMsgPayload;
   #Received_Msg_Status:=#LMQTT_DB.receivedMsgStatus;
   #Received_Msg_Length := #LMQTT_DB.receivedMsgDataLen;
   #LMQTT_DB.enable := #Enable;
   // timeOut := "Settings_DB".Shuttle_MQTT_Settings.Timeout,
   #LMQTT_DB.qos := "Settings_DB".Shuttle_MQTT.QoS;
   #LMQTT_DB.retain := "Settings_DB".Shuttle_MQTT.Retain;
   #Status := #LMQTT_DB.status;

   IF NOT #bSubscribed THEN
       FOR #Shuttle_No := 1 TO "Settings_DB".System.Shuttle_Count DO
           #iIndex := #Shuttle_No;
           #sIndexStr := "RemovePlusSign"(UINT_TO_STRING(#iIndex));
           // preparing names of Topics for subscribing
           #sSubTopic[#Shuttle_No] := CONCAT(IN1 := 'vehicle/', IN2 := 'Shuttle-');
           IF #iIndex < 10 THEN
               #sSubTopic[#Shuttle_No] := CONCAT(IN1 := #sSubTopic[#Shuttle_No], IN2 := '0');
           END_IF;
           #sSubTopic[#Shuttle_No] := CONCAT(IN1 := #sSubTopic[#Shuttle_No], IN2 := #sIndexStr);
           #sSubTopic[#Shuttle_No] := CONCAT(IN1 := #sSubTopic[#Shuttle_No], IN2 := '/state');
       END_FOR;

       #SubscribeCount := 1;
       FOR #Y := 1 TO "Settings_DB".System.Shuttle_Count DO //1-24
           #SubscribeTopicList[#SubscribeCount] := #sSubTopic[#Y];
           IF #Y < "Settings_DB".System.Shuttle_Count THEN
               #SubscribeCount := #SubscribeCount + 1;
           END_IF;
       END_FOR;

       CASE #SubscribeState OF
           0: // Início
               IF #SubscribeIndex <= #SubscribeCount THEN
                   #LMQTT_DB.mqttTopic := STRING_TO_WSTRING(#SubscribeTopicList[#SubscribeIndex]);
                   #LMQTT_DB.subscribe := TRUE; // comando por 1 ciclo
                   #SubscribeState := 1;
               ELSE
                   #SubscribeState := 99; // Tudo assinado
               END_IF;

           1: // Espera pelo DONE
               IF #LMQTT_DB.done THEN
                   #LMQTT_DB.subscribe := FALSE;
                   #SubscribeIndex := #SubscribeIndex + 1;
                   #SubscribeState := 0;
               ELSIF NOT #LMQTT_DB.done AND NOT #LMQTT_DB.subscribe THEN
                   #SubscribeState := 0;
               ELSIF #LMQTT_DB.error THEN
                   // Lidar com erro
                   #SubscribeState := 98;
                   "Error_Word_1".%X2 := TRUE; //MQTT State in Error
               END_IF;

           98: // Erro
               #LMQTT_DB.subscribe := FALSE;
               #bSubscribed := FALSE;

               IF "Reset_All" THEN
                   #SubscribeCount := 0;
                   #SubscribeIndex := 1;
                   #SubscribeState := 0;
                   "Error_Word_1".%X2 := FALSE;
               END_IF;

           99: // Fim
               #bSubscribed := TRUE;
               #LMQTT_DB.subscribe := FALSE;
       END_CASE;
   END_IF;

   FOR #k := 1 TO "Settings_DB".System.Shuttle_Count DO
       IF #LMQTT_DB.receivedTopic = STRING_TO_WSTRING(#sSubTopic[#k]) THEN
           #sPayloadRcv := "ByteArrayToString"(ByteArray := #LMQTT_DB.receivedMsgPayload,
                                               Lenght := UDINT_TO_INT(#LMQTT_DB.receivedMsgDataLen),
                                               ByteArrayToString_1 => #sPayloadRcv_1,
                                               ByteArrayToString_2=>#sPayloadRcv_2,
                                               ByteArrayToString_3=>#sPayloadRcv_3,
                                               ByteArrayToString_4=>#sPayloadRcv_4,
                                               ByteArrayToString_5=>#sPayloadRcv_5);

           IF #sPayloadRcv <> '' THEN
               "Shuttle_MQTT_DB".Shuttle_MQTT[#k].Message.Shuttle_Status := "ParseShuttle_Status"(String_1 := #sPayloadRcv,
                                                                                             String_2 := #sPayloadRcv_1,
                                                                                             String_3 := #sPayloadRcv_2,
                                                                                             String_4:=#sPayloadRcv_3,
                                                                                             String_5:=#sPayloadRcv_4,
                                                                                             String_6:=#sPayloadRcv_5);
           END_IF;
      END_IF;
   END_FOR;


   REGION Cyclic Error Checks

       IF #Error THEN
           //16#8001 Simultaneous input (rising edge) at publish/subscribe/unsubscribe inputs
           IF #Status = 16#8001 THEN
               #Error := 0; // 36:1 
           //16#8200 Client identifier is empty – Client identifier must be at least 1 character long
           ELSIF #Status = 16#8200 THEN
               #Error := 0; // 36:2 
           //16#8201 Broker's hostname OR IP address is invalid
           ELSIF #Status = 16#8201 THEN
               #Error := 0; // 36:3
           //16#8210 Invalid array size:
           //• During connection establishment: Invalid array size at The "willMsgLen" parameter
           //• During publish: Invalid array size at The "publishMsgLen" parameter
           ELSIF #Status = 16#8210 THEN
               #Error := 0; // 36:4
           //16#8220 Invalid value at The "keepAlive" parameter
           ELSIF #Status = 16#8220 THEN
               #Error := 0; // 36:5
           //16#8230 Invalid value at parameter "qos"
           ELSIF #Status = 16#8230 THEN
               #Error := 0; // 36:6
           //16#8300 Topic empty OR invalid (publish)
           ELSIF #Status = 16#8300 THEN
               #Error := 0; // 36:7
           //16#8310 Topic empty OR invalid (subscribe)
           ELSIF #Status = 16#8310 THEN
               #Error := 0; // 36:8
           //16#8320 Topic empty OR invalid (unsubscribe)
           ELSIF #Status = 16#8320 THEN
               #Error := 0; // 36:9
           //16#8600 Undefined state in The state machine
           ELSIF #Status = 16#8600 THEN
               #Error := 0; // 36:10
           //16#8601 #Error OF subordinate instruction "TCON"
           //The #Error code OF The instruction is output at "diagnostics.subfunctionStatus". The meaning OF The respective
           //#Error code can be found in The TIA Portal Information System.
           ELSIF #Status = 16#8601 THEN
               #Error := 0; // 36:60
           //16#8620 connection establishment timeout. IF necessary, increase the "timeOut" value.
           ELSIF #Status = 16#8620 THEN
               #Error := 0; // 36:11
           //16#8650 timeout during The processing OF The job
           ELSIF #Status = 16#8650 THEN
               #Error := 0; // 36:12
           //16#8670 timeout during MQTT connection setup with The MQTT broker
           ELSIF #Status = 16#8670 THEN
               #Error := 0; // 36:13
           //16#8700 Invalid length in received MQTT packet; new connection required
           ELSIF #Status = 16#8700 THEN
               #Error := 0; // 36:14
           //16#8710 Invalid QoS in received MQTT packet; new connection required
           ELSIF #Status = 16#8710 THEN
               #Error := 0; // 36:15
           //16#8720 Existing session at the MQTT broker; new connection required
           ELSIF #Status = 16#8720 THEN
               #Error := 0; // 36:16
           ELSE
               ;
           END_IF;
       END_IF;
   END_REGION

   //Reset the MQTT communication when pressing the reset button
   IF "Reset_All" THEN
       #SubscribeCount := 0;
       #SubscribeIndex := 1;
       #SubscribeState := 0;
       #bSubscribed := FALSE;
   END_IF;

   // AUTO RESET
   IF "LMQTT_DB".enable AND NOT "LMQTT_DB".valid AND NOT "LMQTT_DB".done AND NOT "LMQTT_DB".busy AND "LMQTT_DB".error THEN
       #Enable_AutoReset := TRUE;
   ELSE
       #Enable_AutoReset := FALSE;
       #MQTT_AutoReset := 0;
       "R_Reset_All_False"(CLK:=TRUE);
       IF "R_Reset_All_False".Q THEN
           "Reset_All" := FALSE;
       END_IF;
   END_IF;

   IF #Enable_AutoReset THEN
       CASE #MQTT_AutoReset OF
           0: // Disable MQTT
               #MQTT_AutoReset := #MQTT_AutoReset + 1;
           1: // Disable MQTT
               "LMQTT_DB".enable := FALSE;
               #MQTT_AutoReset := #MQTT_AutoReset + 1;
           2:  // Reset all
               "Reset_All" := TRUE;
               #MQTT_AutoReset := #MQTT_AutoReset + 1;
           3:  // Wait 10 seconds
               #T_AutoReset(IN:=TRUE,
                            PT:=t#10s);
               IF #T_AutoReset.Q THEN
                   #T_AutoReset(IN := FALSE,
                                PT := t#0s);
                                "Reset_All" := FALSE;
                   #MQTT_AutoReset := #MQTT_AutoReset + 1;
               END_IF;

           4:  // Enable again
               "LMQTT_DB".enable := TRUE;
               #MQTT_AutoReset := #MQTT_AutoReset + 1;

           5: //Check or retry
               IF "LMQTT_DB".enable AND NOT "LMQTT_DB".valid AND NOT "LMQTT_DB".done AND NOT "LMQTT_DB".busy AND "LMQTT_DB".error THEN
                   #T_AutoReset(IN := TRUE,
                                PT := t#3s);

                   IF #T_AutoReset.Q THEN
                       #MQTT_AutoReset := 1;
                   END_IF;
               END_IF;


       END_CASE;
   END_IF;
END_FUNCTION_BLOCK

